(* IEC 61131-3 sources: plc-st-coding-agent/progress/evidence/f14_v14_remaining_20261113/jobs/custom_minimax-m27 (part 8) *)

(* ---- self-medium-01.candidate_01.st ---- *)
FUNCTION_BLOCK FB
VAR_INPUT
    recipe     : ARRAY[1..8] OF ST_Recipe;
    selSlot    : INT;
    loadCmd    : BOOL;
    running    : BOOL;
END_VAR
VAR_OUTPUT
    valid      : BOOL;
    loadedID   : INT;
END_VAR
VAR
    prev_loadCmd  : BOOL := FALSE;
    prev_running  : BOOL := FALSE;
    prev_valid    : BOOL := FALSE;
    prev_loadedID : INT  := 0;
    tmp_risingEdge: BOOL;
    tmp_loadOK    : BOOL;
    tmp_recipeValid: BOOL;
END_VAR
VAR_TEMP
    tmp_slotIdx : INT;
END_VAR
// ----------------------------------------------------------------------
// ENGINEERING_CONTRACT
// Outputs & scan-lifetime behavior (cite PUB IDs):
//   valid    : combinational output; activation on rising loadCmd when NOT running;
//              retention (no recalc) while running; no explicit reset.
//   loadedID : stored on successful load (PUB006); retained while running (PUB016);
//              explicit reset to 0 on invalid load or out-of-bounds slot (PUB005).
// Same-scan priority: running > slot-bounds > recipe validation > ratio > temperature.
// Units: ratio in % (99.0..101.0), temperature in °C (30.0..180.0).
// ----------------------------------------------------------------------

// Rising-edge detection for loadCmd
tmp_risingEdge := loadCmd AND NOT prev_loadCmd;

// Slot index captured once per scan to avoid repeated evaluation
tmp_slotIdx := selSlot;

// Compute load-OK guard: rising edge, not running, slot in [1..8]
// Prevents out-of-bounds array access (PUB002, PUB004, PUB005)
tmp_loadOK := tmp_risingEdge AND (NOT running)
              AND (tmp_slotIdx >= 1) AND (tmp_slotIdx <= 8);

IF tmp_loadOK THEN
    // Combine all three validation conditions (PUB003, PUB006, PUB007)
    // recipeID <> 0  -> slot non-empty
    // totalRatio in [99.0, 101.0]
    // temperature in [30.0, 180.0]
    tmp_recipeValid := (recipe[tmp_slotIdx].recipeID <> 0)
                       AND (recipe[tmp_slotIdx].totalRatio >= 99.0)
                       AND (recipe[tmp_slotIdx].totalRatio <= 101.0)
                       AND (recipe[tmp_slotIdx].temperature >= 30.0)
                       AND (recipe[tmp_slotIdx].temperature <= 180.0);

    IF tmp_recipeValid THEN
        loadedID := recipe[tmp_slotIdx].recipeID;
        valid    := TRUE;
    ELSE
        loadedID := 0;
        valid    := FALSE;
    END_IF;
ELSE
    // running=TRUE: ignore load command, hold previous loadedID (PUB016)
    // no rising edge: hold previous outputs (N10-S9)
    loadedID := prev_loadedID;
    valid    := prev_valid;
END_IF;

// Update state for next scan
prev_loadCmd  := loadCmd;
prev_running  := running;
prev_valid    := valid;
prev_loadedID := loadedID;
END_FUNCTION_BLOCK
(* CONTRACT_RULES [{"kind":"hold_until_reset","output":"loadedID","set_input":"loadCmd","reset_input":null}] *)

(* ---- self-medium-01.candidate_02.st ---- *)
TYPE ST_Recipe : STRUCT
    recipeID    : INT;
    totalRatio  : REAL;
    temperature : REAL;
END_STRUCT
END_TYPE;

FUNCTION_BLOCK FB
VAR_INPUT
    recipe     : ARRAY[1..8] OF ST_Recipe;
    selSlot    : INT;
    loadCmd    : BOOL;
    running    : BOOL;
END_VAR
VAR_OUTPUT
    valid      : BOOL;
    loadedID   : INT;
END_VAR
VAR
    prev_loadCmd  : BOOL := FALSE;
    prev_running  : BOOL := FALSE;
    prev_valid    : BOOL := FALSE;
    prev_loadedID : INT  := 0;
    tmp_risingEdge: BOOL;
    tmp_loadOK    : BOOL;
    tmp_recipeValid: BOOL;
END_VAR
VAR_TEMP
    tmp_slotIdx : INT;
END_VAR
// ----------------------------------------------------------------------
// ENGINEERING_CONTRACT
// Outputs & scan-lifetime behavior (cite PUB IDs):
//   valid    : combinational output; activation on rising loadCmd when NOT running;
//              retention (no recalc) while running; no explicit reset.
//   loadedID : stored on successful load (PUB006); retained while running (PUB016);
//              explicit reset to 0 on invalid load or out-of-bounds slot (PUB005).
// Same-scan priority: running > slot-bounds > recipe validation > ratio > temperature.
// Units: ratio in % (99.0..101.0), temperature in °C (30.0..180.0).
// ----------------------------------------------------------------------

// Rising-edge detection for loadCmd
tmp_risingEdge := loadCmd AND NOT prev_loadCmd;

// Slot index captured once per scan to avoid repeated evaluation
tmp_slotIdx := selSlot;

// Compute load-OK guard: rising edge, not running, slot in [1..8]
// Prevents out-of-bounds array access (PUB002, PUB004, PUB005)
tmp_loadOK := tmp_risingEdge AND (NOT running)
              AND (tmp_slotIdx >= 1) AND (tmp_slotIdx <= 8);

IF tmp_loadOK THEN
    // Combine all three validation conditions (PUB003, PUB006, PUB007)
    // recipeID <> 0  -> slot non-empty
    // totalRatio in [99.0, 101.0]
    // temperature in [30.0, 180.0]
    tmp_recipeValid := (recipe[tmp_slotIdx].recipeID <> 0)
                       AND (recipe[tmp_slotIdx].totalRatio >= 99.0)
                       AND (recipe[tmp_slotIdx].totalRatio <= 101.0)
                       AND (recipe[tmp_slotIdx].temperature >= 30.0)
                       AND (recipe[tmp_slotIdx].temperature <= 180.0);

    IF tmp_recipeValid THEN
        loadedID := recipe[tmp_slotIdx].recipeID;
        valid    := TRUE;
    ELSE
        loadedID := 0;
        valid    := FALSE;
    END_IF;
ELSE
    // running=TRUE: ignore load command, hold previous loadedID (PUB016)
    // no rising edge: hold previous outputs (N10-S9)
    loadedID := prev_loadedID;
    valid    := prev_valid;
END_IF;

// Update state for next scan
prev_loadCmd  := loadCmd;
prev_running  := running;
prev_valid    := valid;
prev_loadedID := loadedID;
END_FUNCTION_BLOCK
(* CONTRACT_RULES [{"kind":"hold_until_reset","output":"loadedID","set_input":"loadCmd","reset_input":null}] *)

(* ---- self-medium-01.candidate_03.st ---- *)
TYPE ST_Recipe : STRUCT
    recipeID    : INT;
    totalRatio  : REAL;
    temperature : REAL;
END_STRUCT
END_TYPE;

FUNCTION_BLOCK FB
VAR_INPUT
    recipe     : ARRAY[1..8] OF ST_Recipe;
    selSlot    : INT;
    loadCmd    : BOOL;
    running    : BOOL;
END_VAR
VAR_OUTPUT
    valid      : BOOL;
    loadedID   : INT;
END_VAR
VAR
    prev_loadCmd  : BOOL := FALSE;
    prev_running  : BOOL := FALSE;
    prev_valid    : BOOL := FALSE;
    prev_loadedID : INT  := 0;
    tmp_risingEdge: BOOL;
    tmp_loadOK    : BOOL;
    tmp_recipeValid: BOOL;
END_VAR
VAR_TEMP
    tmp_slotIdx : INT;
END_VAR
// ----------------------------------------------------------------------
// ENGINEERING_CONTRACT
// Outputs & scan-lifetime behavior (cite PUB IDs):
//   valid    : combinational output; activation on rising loadCmd when NOT running;
//              retention (no recalc) while running; no explicit reset.
//   loadedID : stored on successful load (PUB006); retained while running (PUB016);
//              explicit reset to 0 on invalid load or out-of-bounds slot (PUB005).
// Same-scan priority: running > slot-bounds > recipe validation > ratio > temperature.
// Units: ratio in % (99.0..101.0), temperature in °C (30.0..180.0).
// ----------------------------------------------------------------------

// Rising-edge detection for loadCmd
tmp_risingEdge := loadCmd AND NOT prev_loadCmd;

// Slot index captured once per scan to avoid repeated evaluation
tmp_slotIdx := selSlot;

// Compute load-OK guard: rising edge, not running, slot in [1..8]
// Prevents out-of-bounds array access (PUB002, PUB004, PUB005)
tmp_loadOK := tmp_risingEdge AND (NOT running)
              AND (tmp_slotIdx >= 1) AND (tmp_slotIdx <= 8);

IF tmp_loadOK THEN
    // Combine all three validation conditions (PUB003, PUB006, PUB007)
    // recipeID <> 0  -> slot non-empty
    // totalRatio in [99.0, 101.0]
    // temperature in [30.0, 180.0]
    tmp_recipeValid := (recipe[tmp_slotIdx].recipeID <> 0)
                       AND (recipe[tmp_slotIdx].totalRatio >= 99.0)
                       AND (recipe[tmp_slotIdx].totalRatio <= 101.0)
                       AND (recipe[tmp_slotIdx].temperature >= 30.0)
                       AND (recipe[tmp_slotIdx].temperature <= 180.0);

    IF tmp_recipeValid THEN
        loadedID := recipe[tmp_slotIdx].recipeID;
        valid    := TRUE;
    ELSE
        loadedID := 0;
        valid    := FALSE;
    END_IF;
ELSE
    // No rising load edge OR running: hold previous outputs (N10-S9, PUB016)
    // Even when slot is out of bounds, preserve state; no array access needed.
    loadedID := prev_loadedID;
    valid    := prev_valid;
END_IF;

// Explicit out-of-bounds slot guard: rising edge, not running, slot invalid.
// Must NOT touch the array; set valid=FALSE and loadedID=0 per PUB009/PUB043/S5.
IF tmp_risingEdge AND (NOT running) AND ((tmp_slotIdx < 1) OR (tmp_slotIdx > 8)) THEN
    loadedID := 0;
    valid    := FALSE;
END_IF;

// Update state for next scan
prev_loadCmd  := loadCmd;
prev_running  := running;
prev_valid    := valid;
prev_loadedID := loadedID;
END_FUNCTION_BLOCK
(* CONTRACT_RULES [{"kind":"hold_until_reset","output":"loadedID","set_input":"loadCmd","reset_input":null}] *)

(* ---- self-medium-01.patch_base_02.st ---- *)
FUNCTION_BLOCK FB
VAR_INPUT
    recipe     : ARRAY[1..8] OF ST_Recipe;
    selSlot    : INT;
    loadCmd    : BOOL;
    running    : BOOL;
END_VAR
VAR_OUTPUT
    valid      : BOOL;
    loadedID   : INT;
END_VAR
VAR
    prev_loadCmd  : BOOL := FALSE;
    prev_running  : BOOL := FALSE;
    prev_valid    : BOOL := FALSE;
    prev_loadedID : INT  := 0;
    tmp_risingEdge: BOOL;
    tmp_loadOK    : BOOL;
    tmp_recipeValid: BOOL;
END_VAR
VAR_TEMP
    tmp_slotIdx : INT;
END_VAR
// ----------------------------------------------------------------------
// ENGINEERING_CONTRACT
// Outputs & scan-lifetime behavior (cite PUB IDs):
//   valid    : combinational output; activation on rising loadCmd when NOT running;
//              retention (no recalc) while running; no explicit reset.
//   loadedID : stored on successful load (PUB006); retained while running (PUB016);
//              explicit reset to 0 on invalid load or out-of-bounds slot (PUB005).
// Same-scan priority: running > slot-bounds > recipe validation > ratio > temperature.
// Units: ratio in % (99.0..101.0), temperature in °C (30.0..180.0).
// ----------------------------------------------------------------------

// Rising-edge detection for loadCmd
tmp_risingEdge := loadCmd AND NOT prev_loadCmd;

// Slot index captured once per scan to avoid repeated evaluation
tmp_slotIdx := selSlot;

// Compute load-OK guard: rising edge, not running, slot in [1..8]
// Prevents out-of-bounds array access (PUB002, PUB004, PUB005)
tmp_loadOK := tmp_risingEdge AND (NOT running)
              AND (tmp_slotIdx >= 1) AND (tmp_slotIdx <= 8);

IF tmp_loadOK THEN
    // Combine all three validation conditions (PUB003, PUB006, PUB007)
    // recipeID <> 0  -> slot non-empty
    // totalRatio in [99.0, 101.0]
    // temperature in [30.0, 180.0]
    tmp_recipeValid := (recipe[tmp_slotIdx].recipeID <> 0)
                       AND (recipe[tmp_slotIdx].totalRatio >= 99.0)
                       AND (recipe[tmp_slotIdx].totalRatio <= 101.0)
                       AND (recipe[tmp_slotIdx].temperature >= 30.0)
                       AND (recipe[tmp_slotIdx].temperature <= 180.0);

    IF tmp_recipeValid THEN
        loadedID := recipe[tmp_slotIdx].recipeID;
        valid    := TRUE;
    ELSE
        loadedID := 0;
        valid    := FALSE;
    END_IF;
ELSE
    // running=TRUE: ignore load command, hold previous loadedID (PUB016)
    // no rising edge: hold previous outputs (N10-S9)
    loadedID := prev_loadedID;
    valid    := prev_valid;
END_IF;

// Update state for next scan
prev_loadCmd  := loadCmd;
prev_running  := running;
prev_valid    := valid;
prev_loadedID := loadedID;
END_FUNCTION_BLOCK
(* CONTRACT_RULES [{"kind":"hold_until_reset","output":"loadedID","set_input":"loadCmd","reset_input":null}] *)

(* ---- self-medium-01.patch_base_03.st ---- *)
TYPE ST_Recipe : STRUCT
    recipeID    : INT;
    totalRatio  : REAL;
    temperature : REAL;
END_STRUCT
END_TYPE;

FUNCTION_BLOCK FB
VAR_INPUT
    recipe     : ARRAY[1..8] OF ST_Recipe;
    selSlot    : INT;
    loadCmd    : BOOL;
    running    : BOOL;
END_VAR
VAR_OUTPUT
    valid      : BOOL;
    loadedID   : INT;
END_VAR
VAR
    prev_loadCmd  : BOOL := FALSE;
    prev_running  : BOOL := FALSE;
    prev_valid    : BOOL := FALSE;
    prev_loadedID : INT  := 0;
    tmp_risingEdge: BOOL;
    tmp_loadOK    : BOOL;
    tmp_recipeValid: BOOL;
END_VAR
VAR_TEMP
    tmp_slotIdx : INT;
END_VAR
// ----------------------------------------------------------------------
// ENGINEERING_CONTRACT
// Outputs & scan-lifetime behavior (cite PUB IDs):
//   valid    : combinational output; activation on rising loadCmd when NOT running;
//              retention (no recalc) while running; no explicit reset.
//   loadedID : stored on successful load (PUB006); retained while running (PUB016);
//              explicit reset to 0 on invalid load or out-of-bounds slot (PUB005).
// Same-scan priority: running > slot-bounds > recipe validation > ratio > temperature.
// Units: ratio in % (99.0..101.0), temperature in °C (30.0..180.0).
// ----------------------------------------------------------------------

// Rising-edge detection for loadCmd
tmp_risingEdge := loadCmd AND NOT prev_loadCmd;

// Slot index captured once per scan to avoid repeated evaluation
tmp_slotIdx := selSlot;

// Compute load-OK guard: rising edge, not running, slot in [1..8]
// Prevents out-of-bounds array access (PUB002, PUB004, PUB005)
tmp_loadOK := tmp_risingEdge AND (NOT running)
              AND (tmp_slotIdx >= 1) AND (tmp_slotIdx <= 8);

IF tmp_loadOK THEN
    // Combine all three validation conditions (PUB003, PUB006, PUB007)
    // recipeID <> 0  -> slot non-empty
    // totalRatio in [99.0, 101.0]
    // temperature in [30.0, 180.0]
    tmp_recipeValid := (recipe[tmp_slotIdx].recipeID <> 0)
                       AND (recipe[tmp_slotIdx].totalRatio >= 99.0)
                       AND (recipe[tmp_slotIdx].totalRatio <= 101.0)
                       AND (recipe[tmp_slotIdx].temperature >= 30.0)
                       AND (recipe[tmp_slotIdx].temperature <= 180.0);

    IF tmp_recipeValid THEN
        loadedID := recipe[tmp_slotIdx].recipeID;
        valid    := TRUE;
    ELSE
        loadedID := 0;
        valid    := FALSE;
    END_IF;
ELSE
    // running=TRUE: ignore load command, hold previous loadedID (PUB016)
    // no rising edge: hold previous outputs (N10-S9)
    loadedID := prev_loadedID;
    valid    := prev_valid;
END_IF;

// Update state for next scan
prev_loadCmd  := loadCmd;
prev_running  := running;
prev_valid    := valid;
prev_loadedID := loadedID;
END_FUNCTION_BLOCK
(* CONTRACT_RULES [{"kind":"hold_until_reset","output":"loadedID","set_input":"loadCmd","reset_input":null}] *)

(* ---- self-medium-01.raw_candidate_01.st ---- *)
FUNCTION_BLOCK FB
VAR_INPUT
    recipe     : ARRAY[1..8] OF ST_Recipe;
    selSlot    : INT;
    loadCmd    : BOOL;
    running    : BOOL;
END_VAR
VAR_OUTPUT
    valid      : BOOL;
    loadedID   : INT;
END_VAR
VAR
    prev_loadCmd  : BOOL := FALSE;
    prev_running  : BOOL := FALSE;
    prev_valid    : BOOL := FALSE;
    prev_loadedID : INT  := 0;
    tmp_risingEdge: BOOL;
    tmp_loadOK    : BOOL;
    tmp_recipeValid: BOOL;
END_VAR
VAR_TEMP
    tmp_slotIdx : INT;
END_VAR
// ----------------------------------------------------------------------
// ENGINEERING_CONTRACT
// Outputs & scan-lifetime behavior (cite PUB IDs):
//   valid    : combinational output; activation on rising loadCmd when NOT running;
//              retention (no recalc) while running; no explicit reset.
//   loadedID : stored on successful load (PUB006); retained while running (PUB016);
//              explicit reset to 0 on invalid load or out-of-bounds slot (PUB005).
// Same-scan priority: running > slot-bounds > recipe validation > ratio > temperature.
// Units: ratio in % (99.0..101.0), temperature in °C (30.0..180.0).
// ----------------------------------------------------------------------

// Rising-edge detection for loadCmd
tmp_risingEdge := loadCmd AND NOT prev_loadCmd;

// Slot index captured once per scan to avoid repeated evaluation
tmp_slotIdx := selSlot;

// Compute load-OK guard: rising edge, not running, slot in [1..8]
// Prevents out-of-bounds array access (PUB002, PUB004, PUB005)
tmp_loadOK := tmp_risingEdge AND (NOT running)
              AND (tmp_slotIdx >= 1) AND (tmp_slotIdx <= 8);

IF tmp_loadOK THEN
    // Combine all three validation conditions (PUB003, PUB006, PUB007)
    // recipeID <> 0  -> slot non-empty
    // totalRatio in [99.0, 101.0]
    // temperature in [30.0, 180.0]
    tmp_recipeValid := (recipe[tmp_slotIdx].recipeID <> 0)
                       AND (recipe[tmp_slotIdx].totalRatio >= 99.0)
                       AND (recipe[tmp_slotIdx].totalRatio <= 101.0)
                       AND (recipe[tmp_slotIdx].temperature >= 30.0)
                       AND (recipe[tmp_slotIdx].temperature <= 180.0);

    IF tmp_recipeValid THEN
        loadedID := recipe[tmp_slotIdx].recipeID;
        valid    := TRUE;
    ELSE
        loadedID := 0;
        valid    := FALSE;
    END_IF;
ELSE
    // running=TRUE: ignore load command, hold previous loadedID (PUB016)
    // no rising edge: hold previous outputs (N10-S9)
    loadedID := prev_loadedID;
    valid    := prev_valid;
END_IF;

// Update state for next scan
prev_loadCmd  := loadCmd;
prev_running  := running;
prev_valid    := valid;
prev_loadedID := loadedID;
END_FUNCTION_BLOCK
(* CONTRACT_RULES [{"kind":"hold_until_reset","output":"loadedID","set_input":"loadCmd","reset_input":null}] *)

(* ---- self-medium-01.raw_candidate_02.st ---- *)
TYPE ST_Recipe : STRUCT
    recipeID    : INT;
    totalRatio  : REAL;
    temperature : REAL;
END_STRUCT
END_TYPE

FUNCTION_BLOCK FB
VAR_INPUT
    recipe     : ARRAY[1..8] OF ST_Recipe;
    selSlot    : INT;
    loadCmd    : BOOL;
    running    : BOOL;
END_VAR
VAR_OUTPUT
    valid      : BOOL;
    loadedID   : INT;
END_VAR
VAR
    prev_loadCmd  : BOOL := FALSE;
    prev_running  : BOOL := FALSE;
    prev_valid    : BOOL := FALSE;
    prev_loadedID : INT  := 0;
    tmp_risingEdge: BOOL;
    tmp_loadOK    : BOOL;
    tmp_recipeValid: BOOL;
END_VAR
VAR_TEMP
    tmp_slotIdx : INT;
END_VAR
// ----------------------------------------------------------------------
// ENGINEERING_CONTRACT
// Outputs & scan-lifetime behavior (cite PUB IDs):
//   valid    : combinational output; activation on rising loadCmd when NOT running;
//              retention (no recalc) while running; no explicit reset.
//   loadedID : stored on successful load (PUB006); retained while running (PUB016);
//              explicit reset to 0 on invalid load or out-of-bounds slot (PUB005).
// Same-scan priority: running > slot-bounds > recipe validation > ratio > temperature.
// Units: ratio in % (99.0..101.0), temperature in °C (30.0..180.0).
// ----------------------------------------------------------------------

// Rising-edge detection for loadCmd
tmp_risingEdge := loadCmd AND NOT prev_loadCmd;

// Slot index captured once per scan to avoid repeated evaluation
tmp_slotIdx := selSlot;

// Compute load-OK guard: rising edge, not running, slot in [1..8]
// Prevents out-of-bounds array access (PUB002, PUB004, PUB005)
tmp_loadOK := tmp_risingEdge AND (NOT running)
              AND (tmp_slotIdx >= 1) AND (tmp_slotIdx <= 8);

IF tmp_loadOK THEN
    // Combine all three validation conditions (PUB003, PUB006, PUB007)
    // recipeID <> 0  -> slot non-empty
    // totalRatio in [99.0, 101.0]
    // temperature in [30.0, 180.0]
    tmp_recipeValid := (recipe[tmp_slotIdx].recipeID <> 0)
                       AND (recipe[tmp_slotIdx].totalRatio >= 99.0)
                       AND (recipe[tmp_slotIdx].totalRatio <= 101.0)
                       AND (recipe[tmp_slotIdx].temperature >= 30.0)
                       AND (recipe[tmp_slotIdx].temperature <= 180.0);

    IF tmp_recipeValid THEN
        loadedID := recipe[tmp_slotIdx].recipeID;
        valid    := TRUE;
    ELSE
        loadedID := 0;
        valid    := FALSE;
    END_IF;
ELSE
    // running=TRUE: ignore load command, hold previous loadedID (PUB016)
    // no rising edge: hold previous outputs (N10-S9)
    loadedID := prev_loadedID;
    valid    := prev_valid;
END_IF;

// Update state for next scan
prev_loadCmd  := loadCmd;
prev_running  := running;
prev_valid    := valid;
prev_loadedID := loadedID;
END_FUNCTION_BLOCK
(* CONTRACT_RULES [{"kind":"hold_until_reset","output":"loadedID","set_input":"loadCmd","reset_input":null}] *)

(* ---- self-medium-01.raw_candidate_03.st ---- *)
TYPE ST_Recipe : STRUCT
    recipeID    : INT;
    totalRatio  : REAL;
    temperature : REAL;
END_STRUCT
END_TYPE;

FUNCTION_BLOCK FB
VAR_INPUT
    recipe     : ARRAY[1..8] OF ST_Recipe;
    selSlot    : INT;
    loadCmd    : BOOL;
    running    : BOOL;
END_VAR
VAR_OUTPUT
    valid      : BOOL;
    loadedID   : INT;
END_VAR
VAR
    prev_loadCmd  : BOOL := FALSE;
    prev_running  : BOOL := FALSE;
    prev_valid    : BOOL := FALSE;
    prev_loadedID : INT  := 0;
    tmp_risingEdge: BOOL;
    tmp_loadOK    : BOOL;
    tmp_recipeValid: BOOL;
END_VAR
VAR_TEMP
    tmp_slotIdx : INT;
END_VAR
// ----------------------------------------------------------------------
// ENGINEERING_CONTRACT
// Outputs & scan-lifetime behavior (cite PUB IDs):
//   valid    : combinational output; activation on rising loadCmd when NOT running;
//              retention (no recalc) while running; no explicit reset.
//   loadedID : stored on successful load (PUB006); retained while running (PUB016);
//              explicit reset to 0 on invalid load or out-of-bounds slot (PUB005).
// Same-scan priority: running > slot-bounds > recipe validation > ratio > temperature.
// Units: ratio in % (99.0..101.0), temperature in °C (30.0..180.0).
// ----------------------------------------------------------------------

// Rising-edge detection for loadCmd
tmp_risingEdge := loadCmd AND NOT prev_loadCmd;

// Slot index captured once per scan to avoid repeated evaluation
tmp_slotIdx := selSlot;

// Compute load-OK guard: rising edge, not running, slot in [1..8]
// Prevents out-of-bounds array access (PUB002, PUB004, PUB005)
tmp_loadOK := tmp_risingEdge AND (NOT running)
              AND (tmp_slotIdx >= 1) AND (tmp_slotIdx <= 8);

IF tmp_loadOK THEN
    // Combine all three validation conditions (PUB003, PUB006, PUB007)
    // recipeID <> 0  -> slot non-empty
    // totalRatio in [99.0, 101.0]
    // temperature in [30.0, 180.0]
    tmp_recipeValid := (recipe[tmp_slotIdx].recipeID <> 0)
                       AND (recipe[tmp_slotIdx].totalRatio >= 99.0)
                       AND (recipe[tmp_slotIdx].totalRatio <= 101.0)
                       AND (recipe[tmp_slotIdx].temperature >= 30.0)
                       AND (recipe[tmp_slotIdx].temperature <= 180.0);

    IF tmp_recipeValid THEN
        loadedID := recipe[tmp_slotIdx].recipeID;
        valid    := TRUE;
    ELSE
        loadedID := 0;
        valid    := FALSE;
    END_IF;
ELSE
    // No rising load edge OR running: hold previous outputs (N10-S9, PUB016)
    // Even when slot is out of bounds, preserve state; no array access needed.
    loadedID := prev_loadedID;
    valid    := prev_valid;
END_IF;

// Explicit out-of-bounds slot guard: rising edge, not running, slot invalid.
// Must NOT touch the array; set valid=FALSE and loadedID=0 per PUB009/PUB043/S5.
IF tmp_risingEdge AND (NOT running) AND ((tmp_slotIdx < 1) OR (tmp_slotIdx > 8)) THEN
    loadedID := 0;
    valid    := FALSE;
END_IF;

// Update state for next scan
prev_loadCmd  := loadCmd;
prev_running  := running;
prev_valid    := valid;
prev_loadedID := loadedID;
END_FUNCTION_BLOCK
(* CONTRACT_RULES [{"kind":"hold_until_reset","output":"loadedID","set_input":"loadCmd","reset_input":null}] *)

(* ---- self-medium-02.candidate_01.st ---- *)
(* ENGINEERING_CONTRACT: Moving Average Filter (Ring Buffer, 8-point)
 * ---------------------------------------------------------------
 * Input:  enable (BOOL), rawValue (REAL)
 * Output: filteredValue (REAL), windowFull (BOOL), sampleCount (INT)
 *
 * Behavior per output/state:
 *  filteredValue: Combinational arithmetic mean of 1..8 valid samples;
 *                 held unchanged when enable=FALSE (PUB035/S5).
 *                 Units: REAL average of stored REAL samples.
 *  windowFull:    Latch TRUE after sampleCount first reaches 8 (PUB012);
 *                 reset to FALSE on same scan when enable=FALSE (PUB014).
 *                 No explicit reset input; cleared by enable falling edge.
 *  sampleCount:   Monotonic counter 0..8 while enable=TRUE (PUB015/PUB036);
 *                 forced to 0 on same scan when enable=FALSE (PUB014).
 *                 Same-scan priority: clear dominates on enable falling edge.
 *
 * FIFO eviction: When full (count=8), next write overwrites index 1, then 2...
 * First scan (count=0) writes rawValue to index 1; count becomes 1.
 * PUB IDs: PUB001, PUB002, PUB003, PUB004, PUB005, PUB006, PUB007, PUB008,
 *          PUB009, PUB010, PUB011, PUB012, PUB013, PUB014, PUB015, PUB016,
 *          PUB017, PUB018, PUB019, PUB020, PUB021, PUB022, PUB023, PUB024,
 *          PUB025, PUB026, PUB027, PUB028, PUB029, PUB030, PUB031, PUB032,
 *          PUB033, PUB034, PUB035, PUB036, PUB037, PUB038
 *
 * CONTRACT_RULES: [{"kind": "hold_until_reset", "output": "windowFull",
 *                   "set_input": null, "reset_input": "enable"}]
 *)
FUNCTION_BLOCK FB
VAR_INPUT
    enable    : BOOL;
    rawValue  : REAL;
END_VAR
VAR_OUTPUT
    filteredValue : REAL := 0.0;
    windowFull    : BOOL := FALSE;
    sampleCount   : INT  := 0;
END_VAR
VAR
    ringBuffer  : ARRAY[1..8] OF REAL;
    writeIndex  : INT  := 0;
    prev_rawValue : REAL := 0.0;
END_VAR

// Same-scan priority: enable falling edge clears state before any other logic
IF NOT enable THEN
    sampleCount := 0;
    writeIndex  := 0;
    windowFull  := FALSE;
    // filteredValue intentionally NOT written -> retains last value (PUB035)
ELSE
    // enable is TRUE: push sample, compute mean
    writeIndex := ((writeIndex + 1) MOD 8) + 1; // circular 1..8
    ringBuffer[writeIndex] := rawValue;

    IF sampleCount < 8 THEN
        sampleCount := sampleCount + 1;
    END_IF;

    windowFull := (sampleCount = 8); // latch until disable

    // Compute arithmetic mean over actual valid samples only
    VAR i         : INT;
    VAR tmp_sum   : REAL;
    END_VAR
    tmp_sum := 0.0;
    FOR i := 1 TO sampleCount DO
        tmp_sum := tmp_sum + ringBuffer[i];
    END_FOR;
    filteredValue := tmp_sum / TO_REAL(sampleCount);

    prev_rawValue := rawValue;
END_IF;

// Propagate outputs (already assigned in branches above)
END_FUNCTION_BLOCK

(* ---- self-medium-02.candidate_02.st ---- *)
(* ENGINEERING_CONTRACT: Moving Average Filter (Ring Buffer, 8-point)
 * ---------------------------------------------------------------
 * Input:  enable (BOOL), rawValue (REAL)
 * Output: filteredValue (REAL), windowFull (BOOL), sampleCount (INT)
 *
 * Behavior per output/state:
 *  filteredValue: Combinational arithmetic mean of 1..8 valid samples;
 *                 held unchanged when enable=FALSE (PUB035/S5).
 *                 Units: REAL average of stored REAL samples.
 *  windowFull:    Latch TRUE after sampleCount first reaches 8 (PUB012);
 *                 reset to FALSE on same scan when enable=FALSE (PUB014).
 *                 No explicit reset input; cleared by enable falling edge.
 *  sampleCount:   Monotonic counter 0..8 while enable=TRUE (PUB015/PUB036);
 *                 forced to 0 on same scan when enable=FALSE (PUB014).
 *                 Same-scan priority: clear dominates on enable falling edge.
 *
 * FIFO eviction: When full (count=8), next write overwrites index 1, then 2...
 * First scan (count=0) writes rawValue to index 1; count becomes 1.
 * PUB IDs: PUB001, PUB002, PUB003, PUB004, PUB005, PUB006, PUB007, PUB008,
 *          PUB009, PUB010, PUB011, PUB012, PUB013, PUB014, PUB015, PUB016,
 *          PUB017, PUB018, PUB019, PUB020, PUB021, PUB022, PUB023, PUB024,
 *          PUB025, PUB026, PUB027, PUB028, PUB029, PUB030, PUB031, PUB032,
 *          PUB033, PUB034, PUB035, PUB036, PUB037, PUB038
 *
 * CONTRACT_RULES: [{"kind": "hold_until_reset", "output": "windowFull",
 *                   "set_input": null, "reset_input": "enable"}]
 *)
FUNCTION_BLOCK FB
VAR_INPUT
    enable    : BOOL;
    rawValue  : REAL;
END_VAR
VAR_OUTPUT
    filteredValue : REAL := 0.0;
    windowFull    : BOOL := FALSE;
    sampleCount   : INT  := 0;
END_VAR
VAR
    ringBuffer   : ARRAY[1..8] OF REAL;
    writeIndex   : INT  := 0;
    prev_rawValue : REAL := 0.0;
    tmp_i        : INT;
    tmp_sum      : REAL;
END_VAR

// Same-scan priority: enable falling edge clears state before any other logic
IF NOT enable THEN
    sampleCount := 0;
    writeIndex  := 0;
    windowFull  := FALSE;
    // filteredValue intentionally NOT written -> retains last value (PUB035)
ELSE
    // enable is TRUE: push sample, compute mean
    writeIndex := ((writeIndex + 1) MOD 8) + 1; // circular 1..8
    ringBuffer[writeIndex] := rawValue;

    IF sampleCount < 8 THEN
        sampleCount := sampleCount + 1;
    END_IF;

    windowFull := (sampleCount = 8); // latch until disable

    // Compute arithmetic mean over actual valid samples only
    tmp_sum := 0.0;
    FOR tmp_i := 1 TO sampleCount DO
        tmp_sum := tmp_sum + ringBuffer[tmp_i];
    END_FOR;
    filteredValue := tmp_sum / TO_REAL(sampleCount);

    prev_rawValue := rawValue;
END_IF;

// Propagate outputs (already assigned in branches above)
END_FUNCTION_BLOCK

(* ---- self-medium-02.candidate_03.st ---- *)
(* ENGINEERING_CONTRACT: Moving Average Filter (Ring Buffer, 8-point)
 * ---------------------------------------------------------------
 * Input:  enable (BOOL), rawValue (REAL)
 * Output: filteredValue (REAL), windowFull (BOOL), sampleCount (INT)
 *
 * Behavior per output/state:
 *  filteredValue: Combinational arithmetic mean of 1..8 valid samples;
 *                 held unchanged when enable=FALSE (PUB035/S5).
 *                 Units: REAL average of stored REAL samples.
 *  windowFull:    Latch TRUE after sampleCount first reaches 8 (PUB012);
 *                 reset to FALSE on same scan when enable=FALSE (PUB014).
 *                 No explicit reset input; cleared by enable falling edge.
 *  sampleCount:   Monotonic counter 0..8 while enable=TRUE (PUB015/PUB036);
 *                 forced to 0 on same scan when enable=FALSE (PUB014).
 *                 Same-scan priority: clear dominates on enable falling edge.
 *
 * FIFO eviction: When full (count=8), next write overwrites index 1, then 2...
 * First scan (count=0) writes rawValue to index 1; count becomes 1.
 * PUB IDs: PUB001, PUB002, PUB003, PUB004, PUB005, PUB006, PUB007, PUB008,
 *          PUB009, PUB010, PUB011, PUB012, PUB013, PUB014, PUB015, PUB016,
 *          PUB017, PUB018, PUB019, PUB020, PUB021, PUB022, PUB023, PUB024,
 *          PUB025, PUB026, PUB027, PUB028, PUB029, PUB030, PUB031, PUB032,
 *          PUB033, PUB034, PUB035, PUB036, PUB037, PUB038
 *
 * CONTRACT_RULES: [{"kind": "hold_until_reset", "output": "windowFull",
 *                   "set_input": null, "reset_input": "enable"}]
 *)
FUNCTION_BLOCK FB
VAR_INPUT
    enable   : BOOL;
    rawValue : REAL;
END_VAR
VAR_OUTPUT
    filteredValue : REAL := 0.0;
    windowFull    : BOOL := FALSE;
    sampleCount   : INT  := 0;
END_VAR
VAR
    ringBuffer    : ARRAY[1..8] OF REAL;
    writeIndex    : INT  := 0;
    prev_rawValue : REAL := 0.0;
    tmp_i         : INT;
    tmp_sum       : REAL;
END_VAR

// Same-scan priority: enable falling edge clears state before any other logic
IF NOT enable THEN
    sampleCount := 0;
    writeIndex  := 0;
    windowFull  := FALSE;
    // filteredValue intentionally NOT written -> retains last value (PUB035)
ELSE
    // enable is TRUE: push sample, compute mean
    IF sampleCount < 8 THEN
        sampleCount := sampleCount + 1;
        writeIndex  := sampleCount;
    ELSE
        // Buffer full: FIFO eviction, rotate indices 1..7 forward
        FOR tmp_i := 1 TO 7 DO
            ringBuffer[tmp_i] := ringBuffer[tmp_i + 1];
        END_FOR;
        ringBuffer[8] := rawValue;
    END_IF;

    IF sampleCount < 8 THEN
        ringBuffer[sampleCount] := rawValue;
    END_IF;

    windowFull := (sampleCount = 8); // latch until disable

    // Compute arithmetic mean over actual valid samples only
    tmp_sum := 0.0;
    FOR tmp_i := 1 TO sampleCount DO
        tmp_sum := tmp_sum + ringBuffer[tmp_i];
    END_FOR;
    filteredValue := tmp_sum / TO_REAL(sampleCount);

    prev_rawValue := rawValue;
END_IF;

END_FUNCTION_BLOCK

(* ---- self-medium-02.patch_base_02.st ---- *)
(* ENGINEERING_CONTRACT: Moving Average Filter (Ring Buffer, 8-point)
 * ---------------------------------------------------------------
 * Input:  enable (BOOL), rawValue (REAL)
 * Output: filteredValue (REAL), windowFull (BOOL), sampleCount (INT)
 *
 * Behavior per output/state:
 *  filteredValue: Combinational arithmetic mean of 1..8 valid samples;
 *                 held unchanged when enable=FALSE (PUB035/S5).
 *                 Units: REAL average of stored REAL samples.
 *  windowFull:    Latch TRUE after sampleCount first reaches 8 (PUB012);
 *                 reset to FALSE on same scan when enable=FALSE (PUB014).
 *                 No explicit reset input; cleared by enable falling edge.
 *  sampleCount:   Monotonic counter 0..8 while enable=TRUE (PUB015/PUB036);
 *                 forced to 0 on same scan when enable=FALSE (PUB014).
 *                 Same-scan priority: clear dominates on enable falling edge.
 *
 * FIFO eviction: When full (count=8), next write overwrites index 1, then 2...
 * First scan (count=0) writes rawValue to index 1; count becomes 1.
 * PUB IDs: PUB001, PUB002, PUB003, PUB004, PUB005, PUB006, PUB007, PUB008,
 *          PUB009, PUB010, PUB011, PUB012, PUB013, PUB014, PUB015, PUB016,
 *          PUB017, PUB018, PUB019, PUB020, PUB021, PUB022, PUB023, PUB024,
 *          PUB025, PUB026, PUB027, PUB028, PUB029, PUB030, PUB031, PUB032,
 *          PUB033, PUB034, PUB035, PUB036, PUB037, PUB038
 *
 * CONTRACT_RULES: [{"kind": "hold_until_reset", "output": "windowFull",
 *                   "set_input": null, "reset_input": "enable"}]
 *)
FUNCTION_BLOCK FB
VAR_INPUT
    enable    : BOOL;
    rawValue  : REAL;
END_VAR
VAR_OUTPUT
    filteredValue : REAL := 0.0;
    windowFull    : BOOL := FALSE;
    sampleCount   : INT  := 0;
END_VAR
VAR
    ringBuffer  : ARRAY[1..8] OF REAL;
    writeIndex  : INT  := 0;
    prev_rawValue : REAL := 0.0;
END_VAR

// Same-scan priority: enable falling edge clears state before any other logic
IF NOT enable THEN
    sampleCount := 0;
    writeIndex  := 0;
    windowFull  := FALSE;
    // filteredValue intentionally NOT written -> retains last value (PUB035)
ELSE
    // enable is TRUE: push sample, compute mean
    writeIndex := ((writeIndex + 1) MOD 8) + 1; // circular 1..8
    ringBuffer[writeIndex] := rawValue;

    IF sampleCount < 8 THEN
        sampleCount := sampleCount + 1;
    END_IF;

    windowFull := (sampleCount = 8); // latch until disable

    // Compute arithmetic mean over actual valid samples only
    VAR i         : INT;
    VAR tmp_sum   : REAL;
    END_VAR
    tmp_sum := 0.0;
    FOR i := 1 TO sampleCount DO
        tmp_sum := tmp_sum + ringBuffer[i];
    END_FOR;
    filteredValue := tmp_sum / TO_REAL(sampleCount);

    prev_rawValue := rawValue;
END_IF;

// Propagate outputs (already assigned in branches above)
END_FUNCTION_BLOCK

(* ---- self-medium-02.patch_base_03.st ---- *)
(* ENGINEERING_CONTRACT: Moving Average Filter (Ring Buffer, 8-point)
 * ---------------------------------------------------------------
 * Input:  enable (BOOL), rawValue (REAL)
 * Output: filteredValue (REAL), windowFull (BOOL), sampleCount (INT)
 *
 * Behavior per output/state:
 *  filteredValue: Combinational arithmetic mean of 1..8 valid samples;
 *                 held unchanged when enable=FALSE (PUB035/S5).
 *                 Units: REAL average of stored REAL samples.
 *  windowFull:    Latch TRUE after sampleCount first reaches 8 (PUB012);
 *                 reset to FALSE on same scan when enable=FALSE (PUB014).
 *                 No explicit reset input; cleared by enable falling edge.
 *  sampleCount:   Monotonic counter 0..8 while enable=TRUE (PUB015/PUB036);
 *                 forced to 0 on same scan when enable=FALSE (PUB014).
 *                 Same-scan priority: clear dominates on enable falling edge.
 *
 * FIFO eviction: When full (count=8), next write overwrites index 1, then 2...
 * First scan (count=0) writes rawValue to index 1; count becomes 1.
 * PUB IDs: PUB001, PUB002, PUB003, PUB004, PUB005, PUB006, PUB007, PUB008,
 *          PUB009, PUB010, PUB011, PUB012, PUB013, PUB014, PUB015, PUB016,
 *          PUB017, PUB018, PUB019, PUB020, PUB021, PUB022, PUB023, PUB024,
 *          PUB025, PUB026, PUB027, PUB028, PUB029, PUB030, PUB031, PUB032,
 *          PUB033, PUB034, PUB035, PUB036, PUB037, PUB038
 *
 * CONTRACT_RULES: [{"kind": "hold_until_reset", "output": "windowFull",
 *                   "set_input": null, "reset_input": "enable"}]
 *)
FUNCTION_BLOCK FB
VAR_INPUT
    enable    : BOOL;
    rawValue  : REAL;
END_VAR
VAR_OUTPUT
    filteredValue : REAL := 0.0;
    windowFull    : BOOL := FALSE;
    sampleCount   : INT  := 0;
END_VAR
VAR
    ringBuffer   : ARRAY[1..8] OF REAL;
    writeIndex   : INT  := 0;
    prev_rawValue : REAL := 0.0;
    tmp_i        : INT;
    tmp_sum      : REAL;
END_VAR

// Same-scan priority: enable falling edge clears state before any other logic
IF NOT enable THEN
    sampleCount := 0;
    writeIndex  := 0;
    windowFull  := FALSE;
    // filteredValue intentionally NOT written -> retains last value (PUB035)
ELSE
    // enable is TRUE: push sample, compute mean
    writeIndex := ((writeIndex + 1) MOD 8) + 1; // circular 1..8
    ringBuffer[writeIndex] := rawValue;

    IF sampleCount < 8 THEN
        sampleCount := sampleCount + 1;
    END_IF;

    windowFull := (sampleCount = 8); // latch until disable

    // Compute arithmetic mean over actual valid samples only
    tmp_sum := 0.0;
    FOR tmp_i := 1 TO sampleCount DO
        tmp_sum := tmp_sum + ringBuffer[tmp_i];
    END_FOR;
    filteredValue := tmp_sum / TO_REAL(sampleCount);

    prev_rawValue := rawValue;
END_IF;

// Propagate outputs (already assigned in branches above)
END_FUNCTION_BLOCK

(* ---- self-medium-02.patch_base_04.st ---- *)
(* ENGINEERING_CONTRACT: Moving Average Filter (Ring Buffer, 8-point)
 * ---------------------------------------------------------------
 * Input:  enable (BOOL), rawValue (REAL)
 * Output: filteredValue (REAL), windowFull (BOOL), sampleCount (INT)
 *
 * Behavior per output/state:
 *  filteredValue: Combinational arithmetic mean of 1..8 valid samples;
 *                 held unchanged when enable=FALSE (PUB035/S5).
 *                 Units: REAL average of stored REAL samples.
 *  windowFull:    Latch TRUE after sampleCount first reaches 8 (PUB012);
 *                 reset to FALSE on same scan when enable=FALSE (PUB014).
 *                 No explicit reset input; cleared by enable falling edge.
 *  sampleCount:   Monotonic counter 0..8 while enable=TRUE (PUB015/PUB036);
 *                 forced to 0 on same scan when enable=FALSE (PUB014).
 *                 Same-scan priority: clear dominates on enable falling edge.
 *
 * FIFO eviction: When full (count=8), next write overwrites index 1, then 2...
 * First scan (count=0) writes rawValue to index 1; count becomes 1.
 * PUB IDs: PUB001, PUB002, PUB003, PUB004, PUB005, PUB006, PUB007, PUB008,
 *          PUB009, PUB010, PUB011, PUB012, PUB013, PUB014, PUB015, PUB016,
 *          PUB017, PUB018, PUB019, PUB020, PUB021, PUB022, PUB023, PUB024,
 *          PUB025, PUB026, PUB027, PUB028, PUB029, PUB030, PUB031, PUB032,
 *          PUB033, PUB034, PUB035, PUB036, PUB037, PUB038
 *
 * CONTRACT_RULES: [{"kind": "hold_until_reset", "output": "windowFull",
 *                   "set_input": null, "reset_input": "enable"}]
 *)
FUNCTION_BLOCK FB
VAR_INPUT
    enable   : BOOL;
    rawValue : REAL;
END_VAR
VAR_OUTPUT
    filteredValue : REAL := 0.0;
    windowFull    : BOOL := FALSE;
    sampleCount   : INT  := 0;
END_VAR
VAR
    ringBuffer    : ARRAY[1..8] OF REAL;
    writeIndex    : INT  := 0;
    prev_rawValue : REAL := 0.0;
    tmp_i         : INT;
    tmp_sum       : REAL;
END_VAR

// Same-scan priority: enable falling edge clears state before any other logic
IF NOT enable THEN
    sampleCount := 0;
    writeIndex  := 0;
    windowFull  := FALSE;
    // filteredValue intentionally NOT written -> retains last value (PUB035)
ELSE
    // enable is TRUE: push sample, compute mean
    IF sampleCount < 8 THEN
        sampleCount := sampleCount + 1;
        writeIndex  := sampleCount;
    ELSE
        // Buffer full: FIFO eviction, rotate indices 1..7 forward
        FOR tmp_i := 1 TO 7 DO
            ringBuffer[tmp_i] := ringBuffer[tmp_i + 1];
        END_FOR;
        ringBuffer[8] := rawValue;
    END_IF;

    IF sampleCount < 8 THEN
        ringBuffer[sampleCount] := rawValue;
    END_IF;

    windowFull := (sampleCount = 8); // latch until disable

    // Compute arithmetic mean over actual valid samples only
    tmp_sum := 0.0;
    FOR tmp_i := 1 TO sampleCount DO
        tmp_sum := tmp_sum + ringBuffer[tmp_i];
    END_FOR;
    filteredValue := tmp_sum / TO_REAL(sampleCount);

    prev_rawValue := rawValue;
END_IF;

END_FUNCTION_BLOCK

(* ---- self-medium-02.raw_candidate_01.st ---- *)
(* ENGINEERING_CONTRACT: Moving Average Filter (Ring Buffer, 8-point)
 * ---------------------------------------------------------------
 * Input:  enable (BOOL), rawValue (REAL)
 * Output: filteredValue (REAL), windowFull (BOOL), sampleCount (INT)
 *
 * Behavior per output/state:
 *  filteredValue: Combinational arithmetic mean of 1..8 valid samples;
 *                 held unchanged when enable=FALSE (PUB035/S5).
 *                 Units: REAL average of stored REAL samples.
 *  windowFull:    Latch TRUE after sampleCount first reaches 8 (PUB012);
 *                 reset to FALSE on same scan when enable=FALSE (PUB014).
 *                 No explicit reset input; cleared by enable falling edge.
 *  sampleCount:   Monotonic counter 0..8 while enable=TRUE (PUB015/PUB036);
 *                 forced to 0 on same scan when enable=FALSE (PUB014).
 *                 Same-scan priority: clear dominates on enable falling edge.
 *
 * FIFO eviction: When full (count=8), next write overwrites index 1, then 2...
 * First scan (count=0) writes rawValue to index 1; count becomes 1.
 * PUB IDs: PUB001, PUB002, PUB003, PUB004, PUB005, PUB006, PUB007, PUB008,
 *          PUB009, PUB010, PUB011, PUB012, PUB013, PUB014, PUB015, PUB016,
 *          PUB017, PUB018, PUB019, PUB020, PUB021, PUB022, PUB023, PUB024,
 *          PUB025, PUB026, PUB027, PUB028, PUB029, PUB030, PUB031, PUB032,
 *          PUB033, PUB034, PUB035, PUB036, PUB037, PUB038
 *
 * CONTRACT_RULES: [{"kind": "hold_until_reset", "output": "windowFull",
 *                   "set_input": null, "reset_input": "enable"}]
 *)
FUNCTION_BLOCK FB
VAR_INPUT
    enable    : BOOL;
    rawValue  : REAL;
END_VAR
VAR_OUTPUT
    filteredValue : REAL := 0.0;
    windowFull    : BOOL := FALSE;
    sampleCount   : INT  := 0;
END_VAR
VAR
    ringBuffer  : ARRAY[1..8] OF REAL;
    writeIndex  : INT  := 0;
    prev_rawValue : REAL := 0.0;
END_VAR

// Same-scan priority: enable falling edge clears state before any other logic
IF NOT enable THEN
    sampleCount := 0;
    writeIndex  := 0;
    windowFull  := FALSE;
    // filteredValue intentionally NOT written -> retains last value (PUB035)
ELSE
    // enable is TRUE: push sample, compute mean
    writeIndex := ((writeIndex + 1) MOD 8) + 1; // circular 1..8
    ringBuffer[writeIndex] := rawValue;

    IF sampleCount < 8 THEN
        sampleCount := sampleCount + 1;
    END_IF

    windowFull := (sampleCount = 8); // latch until disable

    // Compute arithmetic mean over actual valid samples only
    VAR i         : INT;
    VAR tmp_sum   : REAL;
    END_VAR
    tmp_sum := 0.0;
    FOR i := 1 TO sampleCount DO
        tmp_sum := tmp_sum + ringBuffer[i];
    END_FOR
    filteredValue := tmp_sum / TO_REAL(sampleCount);

    prev_rawValue := rawValue;
END_IF

// Propagate outputs (already assigned in branches above)
END_FUNCTION_BLOCK

(* ---- self-medium-02.raw_candidate_02.st ---- *)
(* ENGINEERING_CONTRACT: Moving Average Filter (Ring Buffer, 8-point)
 * ---------------------------------------------------------------
 * Input:  enable (BOOL), rawValue (REAL)
 * Output: filteredValue (REAL), windowFull (BOOL), sampleCount (INT)
 *
 * Behavior per output/state:
 *  filteredValue: Combinational arithmetic mean of 1..8 valid samples;
 *                 held unchanged when enable=FALSE (PUB035/S5).
 *                 Units: REAL average of stored REAL samples.
 *  windowFull:    Latch TRUE after sampleCount first reaches 8 (PUB012);
 *                 reset to FALSE on same scan when enable=FALSE (PUB014).
 *                 No explicit reset input; cleared by enable falling edge.
 *  sampleCount:   Monotonic counter 0..8 while enable=TRUE (PUB015/PUB036);
 *                 forced to 0 on same scan when enable=FALSE (PUB014).
 *                 Same-scan priority: clear dominates on enable falling edge.
 *
 * FIFO eviction: When full (count=8), next write overwrites index 1, then 2...
 * First scan (count=0) writes rawValue to index 1; count becomes 1.
 * PUB IDs: PUB001, PUB002, PUB003, PUB004, PUB005, PUB006, PUB007, PUB008,
 *          PUB009, PUB010, PUB011, PUB012, PUB013, PUB014, PUB015, PUB016,
 *          PUB017, PUB018, PUB019, PUB020, PUB021, PUB022, PUB023, PUB024,
 *          PUB025, PUB026, PUB027, PUB028, PUB029, PUB030, PUB031, PUB032,
 *          PUB033, PUB034, PUB035, PUB036, PUB037, PUB038
 *
 * CONTRACT_RULES: [{"kind": "hold_until_reset", "output": "windowFull",
 *                   "set_input": null, "reset_input": "enable"}]
 *)
FUNCTION_BLOCK FB
VAR_INPUT
    enable    : BOOL;
    rawValue  : REAL;
END_VAR
VAR_OUTPUT
    filteredValue : REAL := 0.0;
    windowFull    : BOOL := FALSE;
    sampleCount   : INT  := 0;
END_VAR
VAR
    ringBuffer   : ARRAY[1..8] OF REAL;
    writeIndex   : INT  := 0;
    prev_rawValue : REAL := 0.0;
    tmp_i        : INT;
    tmp_sum      : REAL;
END_VAR

// Same-scan priority: enable falling edge clears state before any other logic
IF NOT enable THEN
    sampleCount := 0;
    writeIndex  := 0;
    windowFull  := FALSE;
    // filteredValue intentionally NOT written -> retains last value (PUB035)
ELSE
    // enable is TRUE: push sample, compute mean
    writeIndex := ((writeIndex + 1) MOD 8) + 1; // circular 1..8
    ringBuffer[writeIndex] := rawValue;

    IF sampleCount < 8 THEN
        sampleCount := sampleCount + 1;
    END_IF;

    windowFull := (sampleCount = 8); // latch until disable

    // Compute arithmetic mean over actual valid samples only
    tmp_sum := 0.0;
    FOR tmp_i := 1 TO sampleCount DO
        tmp_sum := tmp_sum + ringBuffer[tmp_i];
    END_FOR;
    filteredValue := tmp_sum / TO_REAL(sampleCount);

    prev_rawValue := rawValue;
END_IF;

// Propagate outputs (already assigned in branches above)
END_FUNCTION_BLOCK

(* ---- self-medium-02.raw_candidate_03.st ---- *)
(* ENGINEERING_CONTRACT: Moving Average Filter (Ring Buffer, 8-point)
 * ---------------------------------------------------------------
 * Input:  enable (BOOL), rawValue (REAL)
 * Output: filteredValue (REAL), windowFull (BOOL), sampleCount (INT)
 *
 * Behavior per output/state:
 *  filteredValue: Combinational arithmetic mean of 1..8 valid samples;
 *                 held unchanged when enable=FALSE (PUB035/S5).
 *                 Units: REAL average of stored REAL samples.
 *  windowFull:    Latch TRUE after sampleCount first reaches 8 (PUB012);
 *                 reset to FALSE on same scan when enable=FALSE (PUB014).
 *                 No explicit reset input; cleared by enable falling edge.
 *  sampleCount:   Monotonic counter 0..8 while enable=TRUE (PUB015/PUB036);
 *                 forced to 0 on same scan when enable=FALSE (PUB014).
 *                 Same-scan priority: clear dominates on enable falling edge.
 *
 * FIFO eviction: When full (count=8), next write overwrites index 1, then 2...
 * First scan (count=0) writes rawValue to index 1; count becomes 1.
 * PUB IDs: PUB001, PUB002, PUB003, PUB004, PUB005, PUB006, PUB007, PUB008,
 *          PUB009, PUB010, PUB011, PUB012, PUB013, PUB014, PUB015, PUB016,
 *          PUB017, PUB018, PUB019, PUB020, PUB021, PUB022, PUB023, PUB024,
 *          PUB025, PUB026, PUB027, PUB028, PUB029, PUB030, PUB031, PUB032,
 *          PUB033, PUB034, PUB035, PUB036, PUB037, PUB038
 *
 * CONTRACT_RULES: [{"kind": "hold_until_reset", "output": "windowFull",
 *                   "set_input": null, "reset_input": "enable"}]
 *)
FUNCTION_BLOCK FB
VAR_INPUT
    enable   : BOOL;
    rawValue : REAL;
END_VAR
VAR_OUTPUT
    filteredValue : REAL := 0.0;
    windowFull    : BOOL := FALSE;
    sampleCount   : INT  := 0;
END_VAR
VAR
    ringBuffer    : ARRAY[1..8] OF REAL;
    writeIndex    : INT  := 0;
    prev_rawValue : REAL := 0.0;
    tmp_i         : INT;
    tmp_sum       : REAL;
END_VAR

// Same-scan priority: enable falling edge clears state before any other logic
IF NOT enable THEN
    sampleCount := 0;
    writeIndex  := 0;
    windowFull  := FALSE;
    // filteredValue intentionally NOT written -> retains last value (PUB035)
ELSE
    // enable is TRUE: push sample, compute mean
    IF sampleCount < 8 THEN
        sampleCount := sampleCount + 1;
        writeIndex  := sampleCount;
    ELSE
        // Buffer full: FIFO eviction, rotate indices 1..7 forward
        FOR tmp_i := 1 TO 7 DO
            ringBuffer[tmp_i] := ringBuffer[tmp_i + 1];
        END_FOR;
        ringBuffer[8] := rawValue;
    END_IF;

    IF sampleCount < 8 THEN
        ringBuffer[sampleCount] := rawValue;
    END_IF;

    windowFull := (sampleCount = 8); // latch until disable

    // Compute arithmetic mean over actual valid samples only
    tmp_sum := 0.0;
    FOR tmp_i := 1 TO sampleCount DO
        tmp_sum := tmp_sum + ringBuffer[tmp_i];
    END_FOR;
    filteredValue := tmp_sum / TO_REAL(sampleCount);

    prev_rawValue := rawValue;
END_IF;

END_FUNCTION_BLOCK

(* ---- self-medium-03.candidate_01.st ---- *)
FUNCTION_BLOCK FB
VAR_INPUT
    openBtn    : BOOL;
    closeBtn   : BOOL;
    openLimit  : BOOL;
    closeLimit : BOOL;
    obstacle   : BOOL;
END_VAR
VAR_OUTPUT
    motorUp    : BOOL;
    motorDown  : BOOL;
    errorFlag  : BOOL;
END_VAR
VAR
    state        : INT;  // 0=IDLE, 1=OPENING, 2=CLOSING, 3=FAULT
    prev_openBtn  : BOOL := FALSE;
    prev_closeBtn : BOOL := FALSE;
END_VAR
VAR_TEMP
    openRising  : BOOL;
    closeRising : BOOL;
    dualRising  : BOOL;
END_VAR
(*
ENGINEERING_CONTRACT
================================================================================
State retention: IDLE/OPENING/CLOSING/FAULT held in state VAR.
Output motorUp: activation on OPENING entry (PUB010), hold until openLimit or
                obstacle or FAULT entry (PUB003/PUB004/PUB012). No reset
                command de-asserts motorUp; only limit/obstacle/FAULT.
Output motorDown: symmetric to motorUp for CLOSING (PUB011).
Output errorFlag: latched hold_until_reset per CONTRACT_RULES, cleared only
                  by dualRising edge with !obstacle (PUB026/PUB036).
Reset priority: obstacle immediate (PUB012), then dualRising reset
                (PUB036), then limit switches (PUB003/PUB004), then idle
                continuation (PUB003). All same-scan; no added delays.
Physical direction rule: motorUp AND motorDown never both TRUE (PUB007).
Units: BOOL scan-synchronous, no timers. Boundary conditions per formal props.
================================================================================
*)
openRising  := openBtn AND NOT prev_openBtn;
closeRising := closeBtn AND NOT prev_closeBtn;
dualRising  := openRising AND closeRising;

motorUp   := FALSE;
motorDown := FALSE;

IF obstacle THEN
    errorFlag := TRUE;
    state     := FAULT;
    RETURN;
END_IF;

CASE state OF
    0: // IDLE
        IF openRising AND NOT closeBtn AND NOT openLimit THEN
            state := OPENING;
            motorUp := TRUE;
        ELSIF closeRising AND NOT openBtn AND NOT closeLimit THEN
            state := CLOSING;
            motorDown := TRUE;
        END_IF;

    1: // OPENING
        IF openLimit THEN
            state := IDLE;
        END_IF;

    2: // CLOSING
        IF closeLimit THEN
            state := IDLE;
        END_IF;

    3: // FAULT
        IF NOT obstacle AND dualRising THEN
            errorFlag := FALSE;
            state     := IDLE;
        ELSE
            errorFlag := TRUE;
        END_IF;
END_CASE;

prev_openBtn  := openBtn;
prev_closeBtn := closeBtn;
END_FUNCTION_BLOCK

(* CONTRACT_RULES [{"kind": "hold_until_reset", "output": "errorFlag", "set_input": "obstacle", "reset_input": "rising(openBtn AND closeBtn)"}] *)

(* ---- self-medium-03.candidate_02.st ---- *)
FUNCTION_BLOCK FB
VAR_INPUT
    openBtn    : BOOL;
    closeBtn   : BOOL;
    openLimit  : BOOL;
    closeLimit : BOOL;
    obstacle   : BOOL;
END_VAR
VAR_OUTPUT
    motorUp    : BOOL;
    motorDown  : BOOL;
    errorFlag  : BOOL;
END_VAR
VAR
    state        : INT;  // 0=IDLE, 1=OPENING, 2=CLOSING, 3=FAULT
    prev_openBtn  : BOOL := FALSE;
    prev_closeBtn : BOOL := FALSE;
END_VAR
VAR_TEMP
    openRising  : BOOL;
    closeRising : BOOL;
    dualRising  : BOOL;
END_VAR
(*
ENGINEERING_CONTRACT
================================================================================
State retention: IDLE/OPENING/CLOSING/FAULT held in state VAR.
Output motorUp: activation on OPENING entry (PUB010), hold until openLimit or
                obstacle or FAULT entry (PUB003/PUB004/PUB012). No reset
                command de-asserts motorUp; only limit/obstacle/FAULT.
Output motorDown: symmetric to motorUp for CLOSING (PUB011).
Output errorFlag: latched hold_until_reset per CONTRACT_RULES, cleared only
                  by dualRising edge with !obstacle (PUB026/PUB036).
Reset priority: obstacle immediate (PUB012), then dualRising reset
                (PUB036), then limit switches (PUB003/PUB004), then idle
                continuation (PUB003). All same-scan; no added delays.
Physical direction rule: motorUp AND motorDown never both TRUE (PUB007).
Units: BOOL scan-synchronous, no timers. Boundary conditions per formal props.
================================================================================
*)
openRising  := openBtn AND NOT prev_openBtn;
closeRising := closeBtn AND NOT prev_closeBtn;
dualRising  := openRising AND closeRising;

motorUp   := FALSE;
motorDown := FALSE;

IF obstacle THEN
    errorFlag := TRUE;
    state     := 3;
    RETURN;
END_IF;

CASE state OF
    0: // IDLE
        IF openRising AND NOT closeBtn AND NOT openLimit THEN
            state := 1;
            motorUp := TRUE;
        ELSIF closeRising AND NOT openBtn AND NOT closeLimit THEN
            state := 2;
            motorDown := TRUE;
        END_IF;

    1: // OPENING
        IF openLimit THEN
            state := 0;
        END_IF;

    2: // CLOSING
        IF closeLimit THEN
            state := 0;
        END_IF;

    3: // FAULT
        IF NOT obstacle AND dualRising THEN
            errorFlag := FALSE;
            state     := 0;
        ELSE
            errorFlag := TRUE;
        END_IF;
END_CASE;

prev_openBtn  := openBtn;
prev_closeBtn := closeBtn;
END_FUNCTION_BLOCK

(* CONTRACT_RULES [{"kind": "hold_until_reset", "output": "errorFlag", "set_input": "obstacle", "reset_input": "rising(openBtn AND closeBtn)"}] *)

(* ---- self-medium-03.candidate_04.st ---- *)
FUNCTION_BLOCK FB
VAR_INPUT
    openBtn    : BOOL;
    closeBtn   : BOOL;
    openLimit  : BOOL;
    closeLimit : BOOL;
    obstacle   : BOOL;
END_VAR
VAR_OUTPUT
    motorUp    : BOOL;
    motorDown  : BOOL;
    errorFlag  : BOOL;
END_VAR
VAR
    state        : INT;  // 0=IDLE, 1=OPENING, 2=CLOSING, 3=FAULT
    prev_openBtn  : BOOL := FALSE;
    prev_closeBtn : BOOL := FALSE;
END_VAR
VAR_TEMP
    openRising  : BOOL;
    closeRising : BOOL;
    dualRising  : BOOL;
END_VAR
(*
ENGINEERING_CONTRACT
================================================================================
State retention: IDLE/OPENING/CLOSING/FAULT held in state VAR.
Output motorUp: activation on OPENING entry (PUB010), hold until openLimit or
                obstacle or FAULT entry (PUB003/PUB004/PUB012). No reset
                command de-asserts motorUp; only limit/obstacle/FAULT.
Output motorDown: symmetric to motorUp for CLOSING (PUB011).
Output errorFlag: latched hold_until_reset per CONTRACT_RULES, cleared only
                  by dualRising edge with !obstacle (PUB026/PUB036).
Reset priority: obstacle immediate (PUB012), then dualRising reset
                (PUB036), then limit switches (PUB003/PUB004), then idle
                continuation (PUB003). All same-scan; no added delays.
Physical direction rule: motorUp AND motorDown never both TRUE (PUB007).
Units: BOOL scan-synchronous, no timers. Boundary conditions per formal props.
================================================================================
*)
openRising  := openBtn AND NOT prev_openBtn;
closeRising := closeBtn AND NOT prev_closeBtn;
dualRising  := openRising AND closeRising;

motorUp   := FALSE;
motorDown := FALSE;

IF obstacle THEN
    errorFlag := TRUE;
    state     := 3;
    RETURN;
END_IF;

CASE state OF
    0: // IDLE
        IF openRising AND NOT closeBtn AND NOT openLimit THEN
            state := 1;
            motorUp := TRUE;
        ELSIF closeRising AND NOT openBtn AND NOT closeLimit THEN
            state := 2;
            motorDown := TRUE;
        END_IF;

    1: // OPENING
        IF openLimit THEN
            state := 0;
        ELSE
            motorUp := TRUE;
        END_IF;

    2: // CLOSING
        IF closeLimit THEN
            state := 0;
        ELSE
            motorDown := TRUE;
        END_IF;

    3: // FAULT
        IF NOT obstacle AND dualRising THEN
            errorFlag := FALSE;
            state     := 0;
        ELSE
            errorFlag := TRUE;
        END_IF;
END_CASE;

prev_openBtn  := openBtn;
prev_closeBtn := closeBtn;
END_FUNCTION_BLOCK

(* CONTRACT_RULES [{"kind": "hold_until_reset", "output": "errorFlag", "set_input": "obstacle", "reset_input": "rising(openBtn AND closeBtn)"}] *)

(* ---- self-medium-03.patch_base_02.st ---- *)
FUNCTION_BLOCK FB
VAR_INPUT
    openBtn    : BOOL;
    closeBtn   : BOOL;
    openLimit  : BOOL;
    closeLimit : BOOL;
    obstacle   : BOOL;
END_VAR
VAR_OUTPUT
    motorUp    : BOOL;
    motorDown  : BOOL;
    errorFlag  : BOOL;
END_VAR
VAR
    state        : INT;  // 0=IDLE, 1=OPENING, 2=CLOSING, 3=FAULT
    prev_openBtn  : BOOL := FALSE;
    prev_closeBtn : BOOL := FALSE;
END_VAR
VAR_TEMP
    openRising  : BOOL;
    closeRising : BOOL;
    dualRising  : BOOL;
END_VAR
(*
ENGINEERING_CONTRACT
================================================================================
State retention: IDLE/OPENING/CLOSING/FAULT held in state VAR.
Output motorUp: activation on OPENING entry (PUB010), hold until openLimit or
                obstacle or FAULT entry (PUB003/PUB004/PUB012). No reset
                command de-asserts motorUp; only limit/obstacle/FAULT.
Output motorDown: symmetric to motorUp for CLOSING (PUB011).
Output errorFlag: latched hold_until_reset per CONTRACT_RULES, cleared only
                  by dualRising edge with !obstacle (PUB026/PUB036).
Reset priority: obstacle immediate (PUB012), then dualRising reset
                (PUB036), then limit switches (PUB003/PUB004), then idle
                continuation (PUB003). All same-scan; no added delays.
Physical direction rule: motorUp AND motorDown never both TRUE (PUB007).
Units: BOOL scan-synchronous, no timers. Boundary conditions per formal props.
================================================================================
*)
openRising  := openBtn AND NOT prev_openBtn;
closeRising := closeBtn AND NOT prev_closeBtn;
dualRising  := openRising AND closeRising;

motorUp   := FALSE;
motorDown := FALSE;

IF obstacle THEN
    errorFlag := TRUE;
    state     := FAULT;
    RETURN;
END_IF;

CASE state OF
    0: // IDLE
        IF openRising AND NOT closeBtn AND NOT openLimit THEN
            state := OPENING;
            motorUp := TRUE;
        ELSIF closeRising AND NOT openBtn AND NOT closeLimit THEN
            state := CLOSING;
            motorDown := TRUE;
        END_IF;

    1: // OPENING
        IF openLimit THEN
            state := IDLE;
        END_IF;

    2: // CLOSING
        IF closeLimit THEN
            state := IDLE;
        END_IF;

    3: // FAULT
        IF NOT obstacle AND dualRising THEN
            errorFlag := FALSE;
            state     := IDLE;
        ELSE
            errorFlag := TRUE;
        END_IF;
END_CASE;

prev_openBtn  := openBtn;
prev_closeBtn := closeBtn;
END_FUNCTION_BLOCK

(* CONTRACT_RULES [{"kind": "hold_until_reset", "output": "errorFlag", "set_input": "obstacle", "reset_input": "rising(openBtn AND closeBtn)"}] *)

(* ---- self-medium-03.patch_base_03.st ---- *)
FUNCTION_BLOCK FB
VAR_INPUT
    openBtn    : BOOL;
    closeBtn   : BOOL;
    openLimit  : BOOL;
    closeLimit : BOOL;
    obstacle   : BOOL;
END_VAR
VAR_OUTPUT
    motorUp    : BOOL;
    motorDown  : BOOL;
    errorFlag  : BOOL;
END_VAR
VAR
    state        : INT;  // 0=IDLE, 1=OPENING, 2=CLOSING, 3=FAULT
    prev_openBtn  : BOOL := FALSE;
    prev_closeBtn : BOOL := FALSE;
END_VAR
VAR_TEMP
    openRising  : BOOL;
    closeRising : BOOL;
    dualRising  : BOOL;
END_VAR
(*
ENGINEERING_CONTRACT
================================================================================
State retention: IDLE/OPENING/CLOSING/FAULT held in state VAR.
Output motorUp: activation on OPENING entry (PUB010), hold until openLimit or
                obstacle or FAULT entry (PUB003/PUB004/PUB012). No reset
                command de-asserts motorUp; only limit/obstacle/FAULT.
Output motorDown: symmetric to motorUp for CLOSING (PUB011).
Output errorFlag: latched hold_until_reset per CONTRACT_RULES, cleared only
                  by dualRising edge with !obstacle (PUB026/PUB036).
Reset priority: obstacle immediate (PUB012), then dualRising reset
                (PUB036), then limit switches (PUB003/PUB004), then idle
                continuation (PUB003). All same-scan; no added delays.
Physical direction rule: motorUp AND motorDown never both TRUE (PUB007).
Units: BOOL scan-synchronous, no timers. Boundary conditions per formal props.
================================================================================
*)
openRising  := openBtn AND NOT prev_openBtn;
closeRising := closeBtn AND NOT prev_closeBtn;
dualRising  := openRising AND closeRising;

motorUp   := FALSE;
motorDown := FALSE;

IF obstacle THEN
    errorFlag := TRUE;
    state     := 3;
    RETURN;
END_IF;

CASE state OF
    0: // IDLE
        IF openRising AND NOT closeBtn AND NOT openLimit THEN
            state := 1;
            motorUp := TRUE;
        ELSIF closeRising AND NOT openBtn AND NOT closeLimit THEN
            state := 2;
            motorDown := TRUE;
        END_IF;

    1: // OPENING
        IF openLimit THEN
            state := 0;
        END_IF;

    2: // CLOSING
        IF closeLimit THEN
            state := 0;
        END_IF;

    3: // FAULT
        IF NOT obstacle AND dualRising THEN
            errorFlag := FALSE;
            state     := 0;
        ELSE
            errorFlag := TRUE;
        END_IF;
END_CASE;

prev_openBtn  := openBtn;
prev_closeBtn := closeBtn;
END_FUNCTION_BLOCK

(* CONTRACT_RULES [{"kind": "hold_until_reset", "output": "errorFlag", "set_input": "obstacle", "reset_input": "rising(openBtn AND closeBtn)"}] *)

(* ---- self-medium-03.patch_base_04.st ---- *)
FUNCTION_BLOCK FB
VAR_INPUT
    openBtn    : BOOL;
    closeBtn   : BOOL;
    openLimit  : BOOL;
    closeLimit : BOOL;
    obstacle   : BOOL;
END_VAR
VAR_OUTPUT
    motorUp    : BOOL;
    motorDown  : BOOL;
    errorFlag  : BOOL;
END_VAR
VAR
    state        : INT;  // 0=IDLE, 1=OPENING, 2=CLOSING, 3=FAULT
    prev_openBtn  : BOOL := FALSE;
    prev_closeBtn : BOOL := FALSE;
END_VAR
VAR_TEMP
    openRising  : BOOL;
    closeRising : BOOL;
    dualRising  : BOOL;
END_VAR
(*
ENGINEERING_CONTRACT
================================================================================
State retention: IDLE/OPENING/CLOSING/FAULT held in state VAR.
Output motorUp: activation on OPENING entry (PUB010), hold until openLimit or
                obstacle or FAULT entry (PUB003/PUB004/PUB012). No reset
                command de-asserts motorUp; only limit/obstacle/FAULT.
Output motorDown: symmetric to motorUp for CLOSING (PUB011).
Output errorFlag: latched hold_until_reset per CONTRACT_RULES, cleared only
                  by dualRising edge with !obstacle (PUB026/PUB036).
Reset priority: obstacle immediate (PUB012), then dualRising reset
                (PUB036), then limit switches (PUB003/PUB004), then idle
                continuation (PUB003). All same-scan; no added delays.
Physical direction rule: motorUp AND motorDown never both TRUE (PUB007).
Units: BOOL scan-synchronous, no timers. Boundary conditions per formal props.
================================================================================
*)
openRising  := openBtn AND NOT prev_openBtn;
closeRising := closeBtn AND NOT prev_closeBtn;
dualRising  := openRising AND closeRising;

motorUp   := FALSE;
motorDown := FALSE;

IF obstacle THEN
    errorFlag := TRUE;
    state     := 3;
    RETURN;
END_IF;

CASE state OF
    0: // IDLE
        IF openRising AND NOT closeBtn AND NOT openLimit THEN
            state := 1;
            motorUp := TRUE;
        ELSIF closeRising AND NOT openBtn AND NOT closeLimit THEN
            state := 2;
            motorDown := TRUE;
        END_IF;

    1: // OPENING
        IF openLimit THEN
            state := 0;
        END_IF;

    2: // CLOSING
        IF closeLimit THEN
            state := 0;
        END_IF;

    3: // FAULT
        IF NOT obstacle AND dualRising THEN
            errorFlag := FALSE;
            state     := 0;
        ELSE
            errorFlag := TRUE;
        END_IF;
END_CASE;

prev_openBtn  := openBtn;
prev_closeBtn := closeBtn;
END_FUNCTION_BLOCK

(* CONTRACT_RULES [{"kind": "hold_until_reset", "output": "errorFlag", "set_input": "obstacle", "reset_input": "rising(openBtn AND closeBtn)"}] *)

(* ---- self-medium-03.raw_candidate_01.st ---- *)
FUNCTION_BLOCK FB
VAR_INPUT
    openBtn    : BOOL;
    closeBtn   : BOOL;
    openLimit  : BOOL;
    closeLimit : BOOL;
    obstacle   : BOOL;
END_VAR
VAR_OUTPUT
    motorUp    : BOOL;
    motorDown  : BOOL;
    errorFlag  : BOOL;
END_VAR
VAR
    state        : INT;  // 0=IDLE, 1=OPENING, 2=CLOSING, 3=FAULT
    prev_openBtn  : BOOL := FALSE;
    prev_closeBtn : BOOL := FALSE;
END_VAR
VAR_TEMP
    openRising  : BOOL;
    closeRising : BOOL;
    dualRising  : BOOL;
END_VAR
(*
ENGINEERING_CONTRACT
================================================================================
State retention: IDLE/OPENING/CLOSING/FAULT held in state VAR.
Output motorUp: activation on OPENING entry (PUB010), hold until openLimit or
                obstacle or FAULT entry (PUB003/PUB004/PUB012). No reset
                command de-asserts motorUp; only limit/obstacle/FAULT.
Output motorDown: symmetric to motorUp for CLOSING (PUB011).
Output errorFlag: latched hold_until_reset per CONTRACT_RULES, cleared only
                  by dualRising edge with !obstacle (PUB026/PUB036).
Reset priority: obstacle immediate (PUB012), then dualRising reset
                (PUB036), then limit switches (PUB003/PUB004), then idle
                continuation (PUB003). All same-scan; no added delays.
Physical direction rule: motorUp AND motorDown never both TRUE (PUB007).
Units: BOOL scan-synchronous, no timers. Boundary conditions per formal props.
================================================================================
*)
openRising  := openBtn AND NOT prev_openBtn;
closeRising := closeBtn AND NOT prev_closeBtn;
dualRising  := openRising AND closeRising;

motorUp   := FALSE;
motorDown := FALSE;

IF obstacle THEN
    errorFlag := TRUE;
    state     := FAULT;
    RETURN;
END_IF;

CASE state OF
    0: // IDLE
        IF openRising AND NOT closeBtn AND NOT openLimit THEN
            state := OPENING;
            motorUp := TRUE;
        ELSIF closeRising AND NOT openBtn AND NOT closeLimit THEN
            state := CLOSING;
            motorDown := TRUE;
        END_IF;

    1: // OPENING
        IF openLimit THEN
            state := IDLE;
        END_IF;

    2: // CLOSING
        IF closeLimit THEN
            state := IDLE;
        END_IF;

    3: // FAULT
        IF NOT obstacle AND dualRising THEN
            errorFlag := FALSE;
            state     := IDLE;
        ELSE
            errorFlag := TRUE;
        END_IF;
END_CASE;

prev_openBtn  := openBtn;
prev_closeBtn := closeBtn;
END_FUNCTION_BLOCK

(* CONTRACT_RULES [{"kind": "hold_until_reset", "output": "errorFlag", "set_input": "obstacle", "reset_input": "rising(openBtn AND closeBtn)"}] *)

(* ---- self-medium-03.raw_candidate_02.st ---- *)
FUNCTION_BLOCK FB
VAR_INPUT
    openBtn    : BOOL;
    closeBtn   : BOOL;
    openLimit  : BOOL;
    closeLimit : BOOL;
    obstacle   : BOOL;
END_VAR
VAR_OUTPUT
    motorUp    : BOOL;
    motorDown  : BOOL;
    errorFlag  : BOOL;
END_VAR
VAR
    state        : INT;  // 0=IDLE, 1=OPENING, 2=CLOSING, 3=FAULT
    prev_openBtn  : BOOL := FALSE;
    prev_closeBtn : BOOL := FALSE;
END_VAR
VAR_TEMP
    openRising  : BOOL;
    closeRising : BOOL;
    dualRising  : BOOL;
END_VAR
(*
ENGINEERING_CONTRACT
================================================================================
State retention: IDLE/OPENING/CLOSING/FAULT held in state VAR.
Output motorUp: activation on OPENING entry (PUB010), hold until openLimit or
                obstacle or FAULT entry (PUB003/PUB004/PUB012). No reset
                command de-asserts motorUp; only limit/obstacle/FAULT.
Output motorDown: symmetric to motorUp for CLOSING (PUB011).
Output errorFlag: latched hold_until_reset per CONTRACT_RULES, cleared only
                  by dualRising edge with !obstacle (PUB026/PUB036).
Reset priority: obstacle immediate (PUB012), then dualRising reset
                (PUB036), then limit switches (PUB003/PUB004), then idle
                continuation (PUB003). All same-scan; no added delays.
Physical direction rule: motorUp AND motorDown never both TRUE (PUB007).
Units: BOOL scan-synchronous, no timers. Boundary conditions per formal props.
================================================================================
*)
openRising  := openBtn AND NOT prev_openBtn;
closeRising := closeBtn AND NOT prev_closeBtn;
dualRising  := openRising AND closeRising;

motorUp   := FALSE;
motorDown := FALSE;

IF obstacle THEN
    errorFlag := TRUE;
    state     := 3;
    RETURN;
END_IF;

CASE state OF
    0: // IDLE
        IF openRising AND NOT closeBtn AND NOT openLimit THEN
            state := 1;
            motorUp := TRUE;
        ELSIF closeRising AND NOT openBtn AND NOT closeLimit THEN
            state := 2;
            motorDown := TRUE;
        END_IF;

    1: // OPENING
        IF openLimit THEN
            state := 0;
        END_IF;

    2: // CLOSING
        IF closeLimit THEN
            state := 0;
        END_IF;

    3: // FAULT
        IF NOT obstacle AND dualRising THEN
            errorFlag := FALSE;
            state     := 0;
        ELSE
            errorFlag := TRUE;
        END_IF;
END_CASE;

prev_openBtn  := openBtn;
prev_closeBtn := closeBtn;
END_FUNCTION_BLOCK

(* CONTRACT_RULES [{"kind": "hold_until_reset", "output": "errorFlag", "set_input": "obstacle", "reset_input": "rising(openBtn AND closeBtn)"}] *)

(* ---- self-medium-03.raw_candidate_04.st ---- *)
FUNCTION_BLOCK FB
VAR_INPUT
    openBtn    : BOOL;
    closeBtn   : BOOL;
    openLimit  : BOOL;
    closeLimit : BOOL;
    obstacle   : BOOL;
END_VAR
VAR_OUTPUT
    motorUp    : BOOL;
    motorDown  : BOOL;
    errorFlag  : BOOL;
END_VAR
VAR
    state        : INT;  // 0=IDLE, 1=OPENING, 2=CLOSING, 3=FAULT
    prev_openBtn  : BOOL := FALSE;
    prev_closeBtn : BOOL := FALSE;
END_VAR
VAR_TEMP
    openRising  : BOOL;
    closeRising : BOOL;
    dualRising  : BOOL;
END_VAR
(*
ENGINEERING_CONTRACT
================================================================================
State retention: IDLE/OPENING/CLOSING/FAULT held in state VAR.
Output motorUp: activation on OPENING entry (PUB010), hold until openLimit or
                obstacle or FAULT entry (PUB003/PUB004/PUB012). No reset
                command de-asserts motorUp; only limit/obstacle/FAULT.
Output motorDown: symmetric to motorUp for CLOSING (PUB011).
Output errorFlag: latched hold_until_reset per CONTRACT_RULES, cleared only
                  by dualRising edge with !obstacle (PUB026/PUB036).
Reset priority: obstacle immediate (PUB012), then dualRising reset
                (PUB036), then limit switches (PUB003/PUB004), then idle
                continuation (PUB003). All same-scan; no added delays.
Physical direction rule: motorUp AND motorDown never both TRUE (PUB007).
Units: BOOL scan-synchronous, no timers. Boundary conditions per formal props.
================================================================================
*)
openRising  := openBtn AND NOT prev_openBtn;
closeRising := closeBtn AND NOT prev_closeBtn;
dualRising  := openRising AND closeRising;

motorUp   := FALSE;
motorDown := FALSE;

IF obstacle THEN
    errorFlag := TRUE;
    state     := 3;
    RETURN;
END_IF;

CASE state OF
    0: // IDLE
        IF openRising AND NOT closeBtn AND NOT openLimit THEN
            state := 1;
            motorUp := TRUE;
        ELSIF closeRising AND NOT openBtn AND NOT closeLimit THEN
            state := 2;
            motorDown := TRUE;
        END_IF;

    1: // OPENING
        IF openLimit THEN
            state := 0;
        ELSE
            motorUp := TRUE;
        END_IF;

    2: // CLOSING
        IF closeLimit THEN
            state := 0;
        ELSE
            motorDown := TRUE;
        END_IF;

    3: // FAULT
        IF NOT obstacle AND dualRising THEN
            errorFlag := FALSE;
            state     := 0;
        ELSE
            errorFlag := TRUE;
        END_IF;
END_CASE;

prev_openBtn  := openBtn;
prev_closeBtn := closeBtn;
END_FUNCTION_BLOCK

(* CONTRACT_RULES [{"kind": "hold_until_reset", "output": "errorFlag", "set_input": "obstacle", "reset_input": "rising(openBtn AND closeBtn)"}] *)

(* ---- self-medium-04.candidate_01.st ---- *)
FUNCTION_BLOCK FB
VAR_INPUT
    startBtn  : BOOL;
    resetBtn  : BOOL;
    doneSensor: BOOL;
    targetVol : REAL;
    flowVol   : REAL;
END_VAR
VAR_OUTPUT
    valveOpen : BOOL;
    fillsToday: INT;
END_VAR
VAR
    state           : INT;        // 0=IDLE, 1=FILLING, 2=PENDING
    prev_startBtn   : BOOL;
    prev_resetBtn   : BOOL;
    prev_valveOpen  : BOOL;
    pendingConfirm  : BOOL;
    accumulatedVol  : REAL;
    rising_startBtn : BOOL;
    rising_resetBtn : BOOL;
    tmp_doConfirm   : BOOL;
END_VAR

// ENGINEERING_CONTRACT
// States: IDLE(0), FILLING(1), PENDING(2)
// Outputs: valveOpen (BOOL, hold open during FILLING until target reached or reset)
//          fillsToday (INT, hold-until-confirm count, saturation at 32767)
// Confirmed fills increment fillsToday by 1 per bottle, cleared on reset
// ResetBtn rising edge (rising_resetBtn) has absolute priority; clears all state
// StartBtn rising edge (rising_startBtn) in IDLE or PENDING starts new bottle
// Confirmation checks doneSensor at valve-close scan; clears pendingConfirm after
// No hidden timers; all state in VAR; explicit edge detection via prev_* vars

(* CONTRACT_RULES [] *)

rising_startBtn := startBtn AND NOT prev_startBtn;
rising_resetBtn := resetBtn  AND NOT prev_resetBtn;

// PUB001: Reset takes priority - ignore everything else this scan
IF rising_resetBtn THEN
    pendingConfirm := FALSE;
    accumulatedVol := 0.0;
    valveOpen      := FALSE;
    fillsToday     := 0;
    prev_startBtn  := startBtn;
    prev_resetBtn  := resetBtn;
    prev_valveOpen := valveOpen;
    RETURN;
END_IF;

// PUB002: Start new bottle when startBtn rises (idle or waiting confirmation)
IF rising_startBtn AND (state = 0 OR state = 2) THEN
    state           := 1;          // FILLING
    pendingConfirm  := FALSE;      // cancel previous pending if any
    accumulatedVol  := flowVol;    // PUB008: start scan counts flow
    IF accumulatedVol >= targetVol THEN
        valveOpen := FALSE;        // PUB014: immediate达标 close
        tmp_doConfirm := doneSensor;
        IF tmp_doConfirm THEN
            IF fillsToday < 32767 THEN
                fillsToday := fillsToday + 1; // PUB030/PUB031: confirm new bottle
            END_IF;
            pendingConfirm := FALSE;
            state := 0;            // back to idle
        ELSE
            pendingConfirm := TRUE;
            state := 2;            // PENDING
        END_IF;
    ELSE
        valveOpen := TRUE;
    END_IF;
    prev_startBtn  := startBtn;
    prev_resetBtn  := resetBtn;
    prev_valveOpen := valveOpen;
    RETURN;
END_IF;

// PUB003: Accumulate flow during filling, including start scan
IF state = 1 THEN
    accumulatedVol := accumulatedVol + flowVol;
    IF accumulatedVol >= targetVol THEN
        valveOpen := FALSE;
        accumulatedVol := targetVol; // PUB035: cap at target
        pendingConfirm := TRUE;
        tmp_doConfirm := doneSensor;
        IF tmp_doConfirm THEN
            // PUB014/PUB004: 本拍关阀后立即确认
            IF fillsToday < 32767 THEN
                fillsToday := fillsToday + 1;
            END_IF;
            pendingConfirm := FALSE;
            state := 0;
        ELSE
            state := 2; // PUB004: wait for future TRUE
        END_IF;
    END_IF;
END_IF;

// PUB004: In PENDING, confirm on first TRUE of doneSensor (unless reset/start)
IF state = 2 AND doneSensor THEN
    IF fillsToday < 32767 THEN
        fillsToday := fillsToday + 1;
    END_IF;
    pendingConfirm := FALSE;
    state := 0;
END_IF;

// PUB047: New start during PENDING cancels pending before start logic
// Handled above by clearing pendingConfirm on rising_startBtn in PENDING

prev_startBtn  := startBtn;
prev_resetBtn  := resetBtn;
prev_valveOpen := valveOpen;
END_FUNCTION_BLOCK

(* ---- self-medium-04.candidate_03.st ---- *)
FUNCTION_BLOCK FB
VAR_INPUT
    startBtn  : BOOL;
    resetBtn  : BOOL;
    doneSensor: BOOL;
    targetVol : REAL;
    flowVol   : REAL;
END_VAR
VAR_OUTPUT
    valveOpen : BOOL;
    fillsToday: INT;
END_VAR
VAR
    state           : INT;        // 0=IDLE, 1=FILLING, 2=PENDING
    prev_startBtn   : BOOL := FALSE;
    prev_resetBtn   : BOOL := FALSE;
    prev_valveOpen  : BOOL := FALSE;
    pendingConfirm  : BOOL;
    accumulatedVol  : REAL := 0.0;
END_VAR

// ENGINEERING_CONTRACT
// States: IDLE(0), FILLING(1), PENDING(2)
// Outputs: valveOpen (BOOL, hold open during FILLING until target reached or reset)
//          fillsToday (INT, hold-until-confirm count, saturation at 32767)
// Confirmed fills increment fillsToday by 1 per bottle, cleared on reset
// ResetBtn rising edge has absolute priority; clears all state and closes valve
// StartBtn rising edge in IDLE or PENDING starts new bottle, cancels pending
// Confirmation checks doneSensor at valve-close scan; clears pendingConfirm after
// No hidden timers; all state in VAR; explicit edge detection via prev_* vars

(* CONTRACT_RULES [] *)

// PUB001: Reset takes priority - ignore everything else this scan
IF resetBtn AND NOT prev_resetBtn THEN
    pendingConfirm := FALSE;
    accumulatedVol := 0.0;
    valveOpen      := FALSE;
    fillsToday     := 0;
    state          := 0;
    prev_startBtn  := resetBtn;
    prev_resetBtn  := resetBtn;
    prev_valveOpen := valveOpen;
    RETURN;
END_IF;

// PUB002/PUB047: Start new bottle when startBtn rises (idle or waiting confirmation)
IF startBtn AND NOT prev_startBtn AND (state = 0 OR state = 2) THEN
    state          := 1;          // FILLING
    pendingConfirm := FALSE;      // cancel previous pending if any
    accumulatedVol := flowVol;    // PUB008: start scan counts flow
    IF accumulatedVol >= targetVol THEN
        valveOpen := FALSE;        // PUB014: immediate达标 close
        IF doneSensor THEN
            IF fillsToday < 32767 THEN
                fillsToday := fillsToday + 1; // PUB030/PUB031: confirm new bottle
            END_IF;
            pendingConfirm := FALSE;
            state := 0;            // back to idle
        ELSE
            pendingConfirm := TRUE;
            state := 2;            // PENDING
        END_IF;
    ELSE
        valveOpen := TRUE;
    END_IF;
    prev_startBtn  := startBtn;
    prev_resetBtn  := resetBtn;
    prev_valveOpen := valveOpen;
    RETURN;
END_IF;

// PUB003: Accumulate flow during filling, including start scan
IF state = 1 THEN
    accumulatedVol := accumulatedVol + flowVol;
    IF accumulatedVol >= targetVol THEN
        valveOpen := FALSE;
        accumulatedVol := targetVol; // PUB035: cap at target
        pendingConfirm := TRUE;
        IF doneSensor THEN
            // PUB014/PUB004: 本拍关阀后立即确认
            IF fillsToday < 32767 THEN
                fillsToday := fillsToday + 1;
            END_IF;
            pendingConfirm := FALSE;
            state := 0;
        ELSE
            state := 2; // PUB004: wait for future TRUE
        END_IF;
    END_IF;
END_IF;

// PUB004: In PENDING, confirm on first TRUE of doneSensor (unless reset/start)
IF state = 2 AND doneSensor THEN
    IF fillsToday < 32767 THEN
        fillsToday := fillsToday + 1;
    END_IF;
    pendingConfirm := FALSE;
    state := 0;
END_IF;

prev_startBtn  := startBtn;
prev_resetBtn  := resetBtn;
prev_valveOpen := valveOpen;
END_FUNCTION_BLOCK

(* ---- self-medium-04.patch_base_02.st ---- *)
FUNCTION_BLOCK FB
VAR_INPUT
    startBtn  : BOOL;
    resetBtn  : BOOL;
    doneSensor: BOOL;
    targetVol : REAL;
    flowVol   : REAL;
END_VAR
VAR_OUTPUT
    valveOpen : BOOL;
    fillsToday: INT;
END_VAR
VAR
    state           : INT;        // 0=IDLE, 1=FILLING, 2=PENDING
    prev_startBtn   : BOOL;
    prev_resetBtn   : BOOL;
    prev_valveOpen  : BOOL;
    pendingConfirm  : BOOL;
    accumulatedVol  : REAL;
    rising_startBtn : BOOL;
    rising_resetBtn : BOOL;
    tmp_doConfirm   : BOOL;
END_VAR

// ENGINEERING_CONTRACT
// States: IDLE(0), FILLING(1), PENDING(2)
// Outputs: valveOpen (BOOL, hold open during FILLING until target reached or reset)
//          fillsToday (INT, hold-until-confirm count, saturation at 32767)
// Confirmed fills increment fillsToday by 1 per bottle, cleared on reset
// ResetBtn rising edge (rising_resetBtn) has absolute priority; clears all state
// StartBtn rising edge (rising_startBtn) in IDLE or PENDING starts new bottle
// Confirmation checks doneSensor at valve-close scan; clears pendingConfirm after
// No hidden timers; all state in VAR; explicit edge detection via prev_* vars

(* CONTRACT_RULES [] *)

rising_startBtn := startBtn AND NOT prev_startBtn;
rising_resetBtn := resetBtn  AND NOT prev_resetBtn;

// PUB001: Reset takes priority - ignore everything else this scan
IF rising_resetBtn THEN
    pendingConfirm := FALSE;
    accumulatedVol := 0.0;
    valveOpen      := FALSE;
    fillsToday     := 0;
    prev_startBtn  := startBtn;
    prev_resetBtn  := resetBtn;
    prev_valveOpen := valveOpen;
    RETURN;
END_IF;

// PUB002: Start new bottle when startBtn rises (idle or waiting confirmation)
IF rising_startBtn AND (state = 0 OR state = 2) THEN
    state           := 1;          // FILLING
    pendingConfirm  := FALSE;      // cancel previous pending if any
    accumulatedVol  := flowVol;    // PUB008: start scan counts flow
    IF accumulatedVol >= targetVol THEN
        valveOpen := FALSE;        // PUB014: immediate达标 close
        tmp_doConfirm := doneSensor;
        IF tmp_doConfirm THEN
            IF fillsToday < 32767 THEN
                fillsToday := fillsToday + 1; // PUB030/PUB031: confirm new bottle
            END_IF;
            pendingConfirm := FALSE;
            state := 0;            // back to idle
        ELSE
            pendingConfirm := TRUE;
            state := 2;            // PENDING
        END_IF;
    ELSE
        valveOpen := TRUE;
    END_IF;
    prev_startBtn  := startBtn;
    prev_resetBtn  := resetBtn;
    prev_valveOpen := valveOpen;
    RETURN;
END_IF;

// PUB003: Accumulate flow during filling, including start scan
IF state = 1 THEN
    accumulatedVol := accumulatedVol + flowVol;
    IF accumulatedVol >= targetVol THEN
        valveOpen := FALSE;
        accumulatedVol := targetVol; // PUB035: cap at target
        pendingConfirm := TRUE;
        tmp_doConfirm := doneSensor;
        IF tmp_doConfirm THEN
            // PUB014/PUB004: 本拍关阀后立即确认
            IF fillsToday < 32767 THEN
                fillsToday := fillsToday + 1;
            END_IF;
            pendingConfirm := FALSE;
            state := 0;
        ELSE
            state := 2; // PUB004: wait for future TRUE
        END_IF;
    END_IF;
END_IF;

// PUB004: In PENDING, confirm on first TRUE of doneSensor (unless reset/start)
IF state = 2 AND doneSensor THEN
    IF fillsToday < 32767 THEN
        fillsToday := fillsToday + 1;
    END_IF;
    pendingConfirm := FALSE;
    state := 0;
END_IF;

// PUB047: New start during PENDING cancels pending before start logic
// Handled above by clearing pendingConfirm on rising_startBtn in PENDING

prev_startBtn  := startBtn;
prev_resetBtn  := resetBtn;
prev_valveOpen := valveOpen;
END_FUNCTION_BLOCK

(* ---- self-medium-04.patch_base_03.st ---- *)
FUNCTION_BLOCK FB
VAR_INPUT
    startBtn  : BOOL;
    resetBtn  : BOOL;
    doneSensor: BOOL;
    targetVol : REAL;
    flowVol   : REAL;
END_VAR
VAR_OUTPUT
    valveOpen : BOOL;
    fillsToday: INT;
END_VAR
VAR
    state           : INT;        // 0=IDLE, 1=FILLING, 2=PENDING
    prev_startBtn   : BOOL;
    prev_resetBtn   : BOOL;
    prev_valveOpen  : BOOL;
    pendingConfirm  : BOOL;
    accumulatedVol  : REAL;
    rising_startBtn : BOOL;
    rising_resetBtn : BOOL;
    tmp_doConfirm   : BOOL;
END_VAR

// ENGINEERING_CONTRACT
// States: IDLE(0), FILLING(1), PENDING(2)
// Outputs: valveOpen (BOOL, hold open during FILLING until target reached or reset)
//          fillsToday (INT, hold-until-confirm count, saturation at 32767)
// Confirmed fills increment fillsToday by 1 per bottle, cleared on reset
// ResetBtn rising edge (rising_resetBtn) has absolute priority; clears all state
// StartBtn rising edge (rising_startBtn) in IDLE or PENDING starts new bottle
// Confirmation checks doneSensor at valve-close scan; clears pendingConfirm after
// No hidden timers; all state in VAR; explicit edge detection via prev_* vars

(* CONTRACT_RULES [] *)

rising_startBtn := startBtn AND NOT prev_startBtn;
rising_resetBtn := resetBtn  AND NOT prev_resetBtn;

// PUB001: Reset takes priority - ignore everything else this scan
IF rising_resetBtn THEN
    pendingConfirm := FALSE;
    accumulatedVol := 0.0;
    valveOpen      := FALSE;
    fillsToday     := 0;
    prev_startBtn  := startBtn;
    prev_resetBtn  := resetBtn;
    prev_valveOpen := valveOpen;
    RETURN;
END_IF;

// PUB002: Start new bottle when startBtn rises (idle or waiting confirmation)
IF rising_startBtn AND (state = 0 OR state = 2) THEN
    state           := 1;          // FILLING
    pendingConfirm  := FALSE;      // cancel previous pending if any
    accumulatedVol  := flowVol;    // PUB008: start scan counts flow
    IF accumulatedVol >= targetVol THEN
        valveOpen := FALSE;        // PUB014: immediate达标 close
        tmp_doConfirm := doneSensor;
        IF tmp_doConfirm THEN
            IF fillsToday < 32767 THEN
                fillsToday := fillsToday + 1; // PUB030/PUB031: confirm new bottle
            END_IF;
            pendingConfirm := FALSE;
            state := 0;            // back to idle
        ELSE
            pendingConfirm := TRUE;
            state := 2;            // PENDING
        END_IF;
    ELSE
        valveOpen := TRUE;
    END_IF;
    prev_startBtn  := startBtn;
    prev_resetBtn  := resetBtn;
    prev_valveOpen := valveOpen;
    RETURN;
END_IF;

// PUB003: Accumulate flow during filling, including start scan
IF state = 1 THEN
    accumulatedVol := accumulatedVol + flowVol;
    IF accumulatedVol >= targetVol THEN
        valveOpen := FALSE;
        accumulatedVol := targetVol; // PUB035: cap at target
        pendingConfirm := TRUE;
        tmp_doConfirm := doneSensor;
        IF tmp_doConfirm THEN
            // PUB014/PUB004: 本拍关阀后立即确认
            IF fillsToday < 32767 THEN
                fillsToday := fillsToday + 1;
            END_IF;
            pendingConfirm := FALSE;
            state := 0;
        ELSE
            state := 2; // PUB004: wait for future TRUE
        END_IF;
    END_IF;
END_IF;

// PUB004: In PENDING, confirm on first TRUE of doneSensor (unless reset/start)
IF state = 2 AND doneSensor THEN
    IF fillsToday < 32767 THEN
        fillsToday := fillsToday + 1;
    END_IF;
    pendingConfirm := FALSE;
    state := 0;
END_IF;

// PUB047: New start during PENDING cancels pending before start logic
// Handled above by clearing pendingConfirm on rising_startBtn in PENDING

prev_startBtn  := startBtn;
prev_resetBtn  := resetBtn;
prev_valveOpen := valveOpen;
END_FUNCTION_BLOCK

(* ---- self-medium-04.patch_base_04.st ---- *)
FUNCTION_BLOCK FB
VAR_INPUT
    startBtn  : BOOL;
    resetBtn  : BOOL;
    doneSensor: BOOL;
    targetVol : REAL;
    flowVol   : REAL;
END_VAR
VAR_OUTPUT
    valveOpen : BOOL;
    fillsToday: INT;
END_VAR
VAR
    state           : INT;        // 0=IDLE, 1=FILLING, 2=PENDING
    prev_startBtn   : BOOL;
    prev_resetBtn   : BOOL;
    prev_valveOpen  : BOOL;
    pendingConfirm  : BOOL;
    accumulatedVol  : REAL;
    rising_startBtn : BOOL;
    rising_resetBtn : BOOL;
    tmp_doConfirm   : BOOL;
END_VAR

// ENGINEERING_CONTRACT
// States: IDLE(0), FILLING(1), PENDING(2)
// Outputs: valveOpen (BOOL, hold open during FILLING until target reached or reset)
//          fillsToday (INT, hold-until-confirm count, saturation at 32767)
// Confirmed fills increment fillsToday by 1 per bottle, cleared on reset
// ResetBtn rising edge (rising_resetBtn) has absolute priority; clears all state
// StartBtn rising edge (rising_startBtn) in IDLE or PENDING starts new bottle
// Confirmation checks doneSensor at valve-close scan; clears pendingConfirm after
// No hidden timers; all state in VAR; explicit edge detection via prev_* vars

(* CONTRACT_RULES [] *)

rising_startBtn := startBtn AND NOT prev_startBtn;
rising_resetBtn := resetBtn  AND NOT prev_resetBtn;

// PUB001: Reset takes priority - ignore everything else this scan
IF rising_resetBtn THEN
    pendingConfirm := FALSE;
    accumulatedVol := 0.0;
    valveOpen      := FALSE;
    fillsToday     := 0;
    prev_startBtn  := startBtn;
    prev_resetBtn  := resetBtn;
    prev_valveOpen := valveOpen;
    RETURN;
END_IF;

// PUB002: Start new bottle when startBtn rises (idle or waiting confirmation)
IF rising_startBtn AND (state = 0 OR state = 2) THEN
    state           := 1;          // FILLING
    pendingConfirm  := FALSE;      // cancel previous pending if any
    accumulatedVol  := flowVol;    // PUB008: start scan counts flow
    IF accumulatedVol >= targetVol THEN
        valveOpen := FALSE;        // PUB014: immediate达标 close
        tmp_doConfirm := doneSensor;
        IF tmp_doConfirm THEN
            IF fillsToday < 32767 THEN
                fillsToday := fillsToday + 1; // PUB030/PUB031: confirm new bottle
            END_IF;
            pendingConfirm := FALSE;
            state := 0;            // back to idle
        ELSE
            pendingConfirm := TRUE;
            state := 2;            // PENDING
        END_IF;
    ELSE
        valveOpen := TRUE;
    END_IF;
    prev_startBtn  := startBtn;
    prev_resetBtn  := resetBtn;
    prev_valveOpen := valveOpen;
    RETURN;
END_IF;

// PUB003: Accumulate flow during filling, including start scan
IF state = 1 THEN
    accumulatedVol := accumulatedVol + flowVol;
    IF accumulatedVol >= targetVol THEN
        valveOpen := FALSE;
        accumulatedVol := targetVol; // PUB035: cap at target
        pendingConfirm := TRUE;
        tmp_doConfirm := doneSensor;
        IF tmp_doConfirm THEN
            // PUB014/PUB004: 本拍关阀后立即确认
            IF fillsToday < 32767 THEN
                fillsToday := fillsToday + 1;
            END_IF;
            pendingConfirm := FALSE;
            state := 0;
        ELSE
            state := 2; // PUB004: wait for future TRUE
        END_IF;
    END_IF;
END_IF;

// PUB004: In PENDING, confirm on first TRUE of doneSensor (unless reset/start)
IF state = 2 AND doneSensor THEN
    IF fillsToday < 32767 THEN
        fillsToday := fillsToday + 1;
    END_IF;
    pendingConfirm := FALSE;
    state := 0;
END_IF;

// PUB047: New start during PENDING cancels pending before start logic
// Handled above by clearing pendingConfirm on rising_startBtn in PENDING

prev_startBtn  := startBtn;
prev_resetBtn  := resetBtn;
prev_valveOpen := valveOpen;
END_FUNCTION_BLOCK
